(* IEC 61131-3 sources: daoli-st-library/DL_Device (part 30) *)

(* ---- FB_DL_SafetyLightCurtainMute.st ---- *)
// FB_DL_SafetyLightCurtainMute v1.0.0
(*==============================================================================
 * 功能描述: C4 安全光栅消隐。双传感器方向判别消隐状态机：eIdle→eArmed→eMuted→
 *           eRestore→eIdle；双模式下行进方向须 S1 先 S2 后（tDirWin 窗内），方向
 *           错误或消隐超窗 tMuteMax 进 eFault 锁存；单模式下光束遮挡直接进入消隐。
 *           bMuteOut 仅在 eMuted 合法窗口励磁——消隐只放行物料方向判别通过，不屏蔽
 *           任何人体进入判别（muted 不等于屏蔽危险），eFault 相 bMuteOut 强制断磁。
 * 接口契约: 输入 bS1/bS2/bDualMode/bMuteReq/tDirWin/tMuteMax/bReset；
 *           输出 bMuteOut/eState/eCause/bError/nErrId。
 * 边界: ① 组态闸：tDirWin<=T#0S、tMuteMax<=T#0S → 故障锁存；② 三枚 R_TRIG + 两枚
 *           TON 段 0 无条件周期刷新；③ 恢复相再次遮挡判超窗违约（安全侧，不续窗）；
 *           ④ 零全局耦合。
 * 码表: 16#0007_0303 故障级总码（组态非法/方向违约/消隐超窗/非法相位，锁存至 bReset
 *       上升沿且光束全清）；16#0007_0403 信息级：消隐窗口有效（励磁中，每拍重算）。
 * 修订历史: 2026-11-23  v1.0.0  R74 首版
 *==============================================================================*)

TYPE E_DL_SlcState :
(
    eIdle    := 0,    // 待命（光束清、无请求）/ Idle, beams clear, no request
    eArmed   := 10,   // 已布防（等待方向判别）/ Armed, awaiting direction discrimination
    eMuted   := 20,   // 消隐励磁中 / Muted, output energised
    eRestore := 30,   // 恢复相（等待光束全清）/ Restore, awaiting beams clear
    eFault   := 90    // 故障锁存相（复位沿 + 光束全清迁出）/ Fault latched
);
END_TYPE

TYPE E_DL_SlcCause :
(
    eNone       := 0,   // 无故障成因 / No cause
    eCfgIllegal := 1,   // 组态非法 / Illegal configuration
    eDirWrong   := 2,   // 方向判别违约（S2 先于 S1）/ Direction violation, S2 before S1
    eMuteOver   := 3,   // 消隐超窗或恢复相再遮挡 / Mute window overrun or re-break in restore
    ePhaseBad   := 4    // 非法相位兜底 / Illegal phase fallback
);
END_TYPE

FUNCTION_BLOCK FB_DL_SafetyLightCurtainMute
VAR_INPUT
    bS1       : BOOL := FALSE;       // 传感器 1（行进侧首束，TRUE=被遮挡）[-] / Sensor 1, entry side, TRUE = blocked
    bS2       : BOOL := FALSE;       // 传感器 2（行进侧次束，TRUE=被遮挡）[-] / Sensor 2, second beam, TRUE = blocked
    bDualMode : BOOL := TRUE;        // 双传感器方向判别模式（FALSE=单传感器）[-] / Dual-sensor direction mode, FALSE = single
    bMuteReq  : BOOL := FALSE;       // 消隐请求（安全控制器电平）[-] / Mute request from safety controller
    tDirWin   : TIME := T#500MS;     // S1→S2 方向判别窗，域 > T#0S [ms] / Direction window, domain > T#0S
    tMuteMax  : TIME := T#10S;       // 消隐最大励磁窗，域 > T#0S [ms] / Maximum mute window, domain > T#0S
    bReset    : BOOL := FALSE;       // 复位，上升沿清故障锁存 [-] / Reset edge clears fault
END_VAR
VAR_OUTPUT
    bMuteOut  : BOOL;                // 消隐励磁输出（仅合法窗口 TRUE）[-] / Mute output, energised in legal window only
    eState    : E_DL_SlcState;       // 状态出口，段尾单点映射 / State outlet
    eCause    : E_DL_SlcCause;       // 故障成因出口（归因唯一） / Fault cause outlet
    bError    : BOOL;                // 故障锁存标志 [-] / Fault latch flag
    nErrId    : UDINT;               // 事件码，0 = 无事件 / Event code, 0 = none
END_VAR
VAR
    _eState  : E_DL_SlcState := E_DL_SlcState.eIdle;   // 内部相位（CASE 唯一写入目标） / Internal phase
    _eCause  : E_DL_SlcCause := E_DL_SlcCause.eNone;   // 故障成因锁存量 / Latched cause
    rtS1     : R_TRIG;               // S1 上升沿实例，段 0 无条件刷新 / S1 rising edge instance
    rtS2     : R_TRIG;               // S2 上升沿实例，段 0 无条件刷新 / S2 rising edge instance
    rtReset  : R_TRIG;               // 复位沿实例，段 0 无条件刷新 / Reset edge instance
    tonDir   : TON;                  // 方向判别窗计时（S1 遮挡期间），段 0 无条件刷新 / Direction window timer
    tonMute  : TON;                  // 消隐励磁窗计时，段 0 无条件刷新 / Mute window timer
    _bCfgBad : BOOL;                 // 组态非法当拍量 [-] / Illegal configuration this scan
    _bFault  : BOOL;                 // 故障锁存位（锁存量） / Latched fault bit
    _uFault  : UDINT;                // 故障码锁存（锁存量） / Latched fault code
    _uInfo   : UDINT;                // 信息码，每拍重算 / Info code, recomputed each scan
    _bClear  : BOOL;                 // 光束全清当拍量 [-] / All beams clear this scan
    _bArmedOk: BOOL;                 // 布防前置成立当拍量 [-] / Arming precondition this scan
END_VAR

(* —— 段 0：沿实例与定时器无条件周期刷新（禁置于 IF/CASE 内） —— *)
rtS1(CLK := bS1);                                                  // S1 沿，每拍必调 / S1 edge every scan
rtS2(CLK := bS2);                                                  // S2 沿，每拍必调 / S2 edge every scan
rtReset(CLK := bReset);                                            // 复位沿，每拍必调 / Reset edge every scan
tonDir(IN := (_eState = E_DL_SlcState.eArmed) AND bS1, PT := tDirWin);    // 方向窗（布防相 S1 遮挡期）/ Direction timer while armed and S1 blocked
tonMute(IN := (_eState = E_DL_SlcState.eMuted), PT := tMuteMax);   // 消隐窗（励磁相独占）/ Mute timer while muted

(* —— 段 1：单拍量预清零（锁存量 _bFault/_uFault/_eCause 不入清单） —— *)
bError := FALSE;                                                   // 故障标志预清（置位处同拍回填） / Error flag preset
bMuteOut := FALSE;                                                 // 励磁输出预清（eMuted 相回填） / Mute output preset
_uInfo := 16#0000_0000;                                            // 信息码每拍重算 / Info recomputed every scan
nErrId := 16#0000_0000;                                            // 事件码缺省无事件 / Event code default none
_bClear := (NOT bS1) AND (NOT bS2);                                // 光束全清当拍量 / Beams clear this scan
_bArmedOk := _bClear AND bMuteReq AND (NOT _bFault);               // 布防前置：光束清 + 请求在 / Arming precondition

(* —— 段 2：组态域闸 —— *)
_bCfgBad := (tDirWin <= T#0S) OR (tMuteMax <= T#0S);               // 时间域闸（防窗口恒成立） / Time domain gates

(* —— 段 3：故障锁存与解除（R45 配对；解除沿 = 复位沿 + 组态合法 + 光束全清） —— *)
IF _bCfgBad THEN                                                   // 组态非法 / Illegal configuration
    _uFault := 16#0007_0303;                                       // 故障级总码 / Fault-level code
    _bFault := TRUE;
    bError  := TRUE;
    _eCause := E_DL_SlcCause.eCfgIllegal;                          // 归因：组态非法 / Cause: illegal configuration
END_IF
IF rtReset.Q AND (NOT _bCfgBad) AND _bClear THEN                   // 解除沿（当拍量，光束全清） / Release edge with beams clear
    _bFault := FALSE;                                              // 清故障锁存 / Clear fault latch
    _uFault := 16#0000_0000;                                       // 清故障码 / Clear fault code
    _eCause := E_DL_SlcCause.eNone;                                // 清成因 / Clear cause
    IF _eState = E_DL_SlcState.eFault THEN
        _eState := E_DL_SlcState.eIdle;                            // 故障相唯一迁出路径 / Sole exit from fault phase
    END_IF
END_IF

(* —— 段 4：相位机（ENUM 全成员显式标签 + ELSE 兜底） —— *)
CASE _eState OF

E_DL_SlcState.eIdle:
    IF _bFault THEN                                                // 出口 1：故障锁存 / Fault latched
        _eState := E_DL_SlcState.eFault;
    ELSIF _bArmedOk THEN                                           // 出口 2：前置成立进布防 / Preconditions met, arm
        _eState := E_DL_SlcState.eArmed;
    END_IF

E_DL_SlcState.eArmed:
    IF _bFault THEN                                                // 出口 1：故障锁存 / Fault latched
        _eState := E_DL_SlcState.eFault;
    ELSIF (NOT bMuteReq) OR _bCfgBad THEN                          // 出口 2：请求撤销或组态坏 → 回待命 / Request dropped, back to idle
        _eState := E_DL_SlcState.eIdle;
    ELSIF bDualMode THEN                                           // 双传感器模式分支 / Dual-sensor branch
        IF rtS2.Q AND (NOT bS1) THEN                               // 方向违约：S2 先遮挡而 S1 未遮挡 / Direction violation, S2 first
            _uFault := 16#0007_0303;
            _bFault := TRUE;
            bError  := TRUE;
            _eCause := E_DL_SlcCause.eDirWrong;                    // 归因：方向违约 / Cause: direction violation
            _eState := E_DL_SlcState.eFault;
        ELSIF rtS2.Q AND bS1 THEN                                  // 合法方向：S1 已遮挡后 S2 到 → 进励磁 / Legal direction, enter muted
            _eState := E_DL_SlcState.eMuted;
        ELSIF tonDir.Q THEN                                        // S1 遮挡超方向窗（判别失败安全退） / S1 blocked over direction window
            _eState := E_DL_SlcState.eIdle;
        END_IF
    ELSE                                                           // 单传感器模式：遮挡即励磁 / Single mode, block enters muted
        IF bS1 THEN
            _eState := E_DL_SlcState.eMuted;
        END_IF
    END_IF

E_DL_SlcState.eMuted:
    IF _bFault THEN                                                // 出口 1：故障锁存 / Fault latched
        _eState := E_DL_SlcState.eFault;
    ELSIF tonMute.Q THEN                                           // 出口 2：励磁超最大窗 → 强制恢复 / Mute window overrun
        _uFault := 16#0007_0303;                                   // 故障级：消隐超窗（超窗不续磁） / Fault, window overrun
        _bFault := TRUE;
        bError  := TRUE;
        _eCause := E_DL_SlcCause.eMuteOver;                        // 归因：超窗 / Cause: window overrun
        _eState := E_DL_SlcState.eRestore;
    ELSIF (NOT bMuteReq) THEN                                      // 出口 3：请求撤销进恢复 / Request dropped, restore
        _eState := E_DL_SlcState.eRestore;
    ELSE
        _uInfo := 16#0007_0403;                                    // 信息级：消隐励磁中 / Info: mute energised
    END_IF

E_DL_SlcState.eRestore:
    IF _bFault THEN                                                // 出口 1：故障锁存 / Fault latched
        _eState := E_DL_SlcState.eFault;
    ELSIF bS1 OR bS2 THEN                                          // 出口 2：恢复相再遮挡 = 违约（不续窗，安全侧） / Re-break in restore, fault
        _uFault := 16#0007_0303;
        _bFault := TRUE;
        bError  := TRUE;
        _eCause := E_DL_SlcCause.eMuteOver;                        // 归因：恢复相再遮挡 / Cause: re-break in restore
        _eState := E_DL_SlcState.eFault;
    ELSE
        _eState := E_DL_SlcState.eIdle;                            // 出口 3：光束全清回待命 / Beams clear, back to idle
    END_IF

E_DL_SlcState.eFault:
    ;                                                              // 故障相：仅段 3 解除沿可迁出（励磁强制断） / Only the release edge leaves, output forced off

ELSE
    _uFault := 16#0007_0303;                                       // 故障级：非法相位兜底 / Illegal-phase fallback
    _bFault := TRUE;
    bError  := TRUE;
    _eCause := E_DL_SlcCause.ePhaseBad;                            // 归因：非法相位 / Cause: illegal phase
    _eState := E_DL_SlcState.eFault;                               // 强拉故障相 / Force fault phase

END_CASE

(* —— 段 5：出口单点映射（名实同源；锁存码回放；故障相励磁强制断） —— *)
IF (_eState = E_DL_SlcState.eMuted) AND (NOT _bFault) THEN
    bMuteOut := TRUE;                                              // 仅合法励磁相输出 / Output only in legal muted phase
END_IF
IF _bFault THEN
    nErrId := _uFault;                                             // 故障锁存码回放 / Replay latched fault code
ELSE
    nErrId := _uInfo;                                              // 信息码 / Info code
END_IF
bError := _bFault;                                                 // 故障标志与锁存同源 / Flag from latch
eState := _eState;                                                 // 状态出口 / State outlet
eCause := _eCause;                                                 // 成因出口 / Cause outlet

END_FUNCTION_BLOCK

(* ---- FB_DL_SafetyRelayFeedback.st ---- *)
(*==============================================================================
 * 组件名称 (Component)  : FB_DL_SafetyRelayFeedback
 * 所属子库 (Sublibrary) : DL_Device
 * 当前版本 (Version)    : 1.0.0
 * 兼容性   (Platform)   : CODESYS 3.5+ / TwinCAT 3 / 汇川 InoProShop / 施耐德 Machine Expert
 *                         仅依赖 Standard.library（TON / R_TRIG）与库内健康枚举唯一属主，
 *                         零厂商私有库
 * 功能描述 (Function)   : 安全继电器（双通道触点）反馈一致性监视。指令 bCmd 变化后开
 *                         tSyncWin 同步窗，窗内应两通道同步跟随；窗末判定四类结局：
 *                         ① 两通道仍不一致 → 通道不同步故障（eSync）；
 *                         ② 仅通道 1 未跟随 → 通道 1 失效（eCh1Fail）；
 *                         ③ 仅通道 2 未跟随 → 通道 2 失效（eCh2Fail）；
 *                         ④ 两通道都未跟随 → 双通道失效（eBothFail）。
 *                         另连续监视常闭回路断开：bNcLogic 为真时「指令为 FALSE 而两通道反馈
 *                         仍为 FALSE」即常闭回路断开（eNcOpen，典型断线/线圈失电）。
 * 安全声明 (Safety)     : **本件不实现任何安全认证功能**。它是反馈一致性监视器，不是安全功能
 *                         的组成部分：不提供双通道自诊断覆盖率证明，不参与 ISO 13849 / IEC 62061
 *                         的 PL / SIL 定级，其输出不得接入安全链路的停机判据。
 * 归属声明 (Ownership)  : 健康出口 eHealth 引用枚举 `E_DL_Ne107Status` 的**唯一属主**，属主文件为
 *                         `C:\Library\DL_Device\I_DL_DeviceHealth.st`（枚举定义位于该文件 L91 附近），
 *                         本件**只引用不重复声明**（全库同名枚举定义计数必须为 1，R67）。
 * 接口     (Interface)  : 输入 bFbCh1 / bFbCh2 双通道反馈、bCmd 指令、tSyncWin 同步窗、bNcLogic
 *                         常闭逻辑组态位、bReset 复位；输出 eCause 归因、bSyncOk 双通道同步、
 *                         eHealth NE107 健康态、eState / bError / nErrId。
 * 边界     (Boundary)   : ① 组态闸：tSyncWin <= T#0S → 故障锁存，**且非法时 eHealth 直接给
 *                         eFailure**（保守：无法判定同步即按失效上报）；
 *                         ② 常闭语义：bNcLogic = TRUE 时期望反馈 = NOT bCmd；= FALSE 时期望 = bCmd；
 *                         ③ 两通道互斥用布尔 XOR 判，无浮点参与；
 *                         ④ TON 两枚 + R_TRIG 两枚段 0 无条件周期刷新（IN 由相位派生，R228A）；
 *                         ⑤ 故障相迁出唯一路径 = bReset 上升沿；⑥ 零全局耦合（无 GVL / 无物理地址）。
 * 解除式   (Release)    : bReset 上升沿 ∧ 组态合法 ∧ 两通道当前一致（bFbCh1 = bFbCh2，当拍量，
 *                         R240 范式）。自证可满足（终审两式 1）：两枚 TON 的 IN 均挂相位，
 *                         故障相内 IN 恒假 → Q 恒假；两通道物理恢复一致即达，无恒假因子。
 * 码表     (Codes)      : 16#0003_0701 故障级：安全继电器反馈故障总码（组态非法 / 通道不同步 /
 *                         单通道失效 / 双通道失效 / 常闭回路断开 / 非法相位），锁存至 bReset 上升沿，
 *                         归因由 eCause 承载（R190 单件单总码，每个成因成员均有独立赋值点）；
 *                         16#0003_0480 信息级：同步窗正常结束（两通道已按指令同步跟随）。
 *                         加码反证（R90）：同步窗正常结束时 bSyncOk 由假转真，而「一直停在 eRun
 *                         未做过切换」也保持 bSyncOk 为真，二者出口组合无法唯一区分「刚完成一次
 *                         动作确认」与「从未动作」，故立一码留痕。
 *                         码段说明：Device 的 03xx 故障子带已占满（03A0~03FF 连续占位，仅余
 *                         03C5~03C9 碎片孔洞），按实战规则 13「禁止回填他人预留碎片孔洞」，
 *                         本批新开 07xx 故障子带并取 16#0003_0701；信息级仍用 04xx 子带取
 *                         16#0003_0480（该段源码实扫为空）。分段理由即此，非笔误。
 * 开源溯源 (Origin)     : 道莅自研 clean-room（参考 ISA-18.2 / NE107 安全回路一致性语义与
 *                         参数域，零代码行复制；t2-8-isa182 族）
 * 修订历史 (Revision)   : 2026-11-19  v1.0.0  R45 首版（批次 3 · 序号 15）
 *==============================================================================*)

TYPE E_DL_SrfState :
(
    eIdle     := 0,     // 未使能待机 / Idle, standing by
    eSyncWait := 10,    // 指令变化后同步窗内（信号暂不可信） / Inside sync window after a command change
    eRun      := 20,    // 同步完成，稳态监视 / Synchronised, steady monitoring
    eFault    := 90     // 故障锁存相 / Fault latched phase
);
END_TYPE

TYPE E_DL_SrfCause :
(
    eNone       := 0,   // 无故障成因 / No cause
    eCfgIllegal := 1,   // 组态非法 / Illegal configuration
    eSync       := 2,   // 两通道不同步 / Channels out of sync
    eCh1Fail    := 3,   // 通道 1 未跟随 / Channel 1 failed to follow
    eCh2Fail    := 4,   // 通道 2 未跟随 / Channel 2 failed to follow
    eBothFail   := 5,   // 两通道均未跟随 / Both channels failed to follow
    eNcOpen     := 6,   // 常闭回路断开 / Normally-closed loop open
    ePhaseBad   := 7    // 非法相位兜底 / Illegal phase fallback
);
END_TYPE

FUNCTION_BLOCK FB_DL_SafetyRelayFeedback
VAR_INPUT
    bFbCh1    : BOOL := FALSE;          // 通道 1 反馈 [-] / Channel 1 feedback
    bFbCh2    : BOOL := FALSE;          // 通道 2 反馈 [-] / Channel 2 feedback
    bCmd      : BOOL := FALSE;          // 继电器指令 [-] / Relay command
    tSyncWin  : TIME := T#300MS;        // 同步窗时长，域 > T#0S [ms] / Sync window duration, domain > T#0S [ms]
    bNcLogic  : BOOL := TRUE;           // 常闭逻辑组态位：TRUE 时期望反馈 = NOT bCmd [-] / NC logic: expected = NOT command
    bReset    : BOOL := FALSE;          // 复位命令，上升沿清故障 [-] / Reset command, rising edge clears fault
END_VAR
VAR_OUTPUT
    eCause    : E_DL_SrfCause;          // 故障成因出口（R190 归因唯一） / Fault cause outlet
    bSyncOk   : BOOL;                   // 双通道同步（稳态且两通道一致且均符合期望） [-] / Channels in sync
    eHealth   : E_DL_Ne107Status;       // NE107 健康态（引用唯一属主枚举） [-] / NE107 health, owner enum referenced
    eState    : E_DL_SrfState;          // 状态出口，段 6 单点映射 / State outlet
    bError    : BOOL;                   // 故障锁存标志 [-] / Fault latch flag
    nErrId    : UDINT;                  // 事件码，0 = 无事件 / Event code, 0 = no event
END_VAR
VAR
    _eState   : E_DL_SrfState := E_DL_SrfState.eIdle;      // 内部相位（CASE 唯一写入目标） / Internal phase
    _eCause   : E_DL_SrfCause := E_DL_SrfCause.eNone;      // 故障成因锁存（锁存量） / Latched cause
    tonSync   : TON;                    // 同步窗计时，段 0 无条件调用 / Sync window timer
    tonDiff   : TON;                    // 通道不一致持续计时，段 0 无条件调用 / Channel-difference timer
    rtCmd     : R_TRIG;                 // 指令变化沿实例，段 0 无条件调用 / Command change edge
    rtReset   : R_TRIG;                 // 复位沿实例，段 0 无条件调用 / Reset edge
    _bExpect  : BOOL;                   // 常闭/常开语义换算后的期望反馈当拍量 [-] / Expected feedback after NC/NO mapping
    _bChDiff  : BOOL;                   // 两通道不一致当拍量 [-] / Channels disagree
    _bCh1Ok   : BOOL;                   // 通道 1 符合期望当拍量 [-] / Channel 1 matches expectation
    _bCh2Ok   : BOOL;                   // 通道 2 符合期望当拍量 [-] / Channel 2 matches expectation
    _bNcOpen  : BOOL;                   // 常闭回路断开当拍量 [-] / NC loop open
    _bCfgBad  : BOOL;                   // 组态非法当拍量 [-] / Illegal configuration
    _bFault   : BOOL;                   // 故障锁存位（锁存量） / Latched fault bit
    _uFault   : UDINT;                  // 故障码锁存（锁存量） / Latched fault code
    _uInfo    : UDINT;                  // 信息码，每拍重算 / Info code, recomputed each scan
END_VAR

(* —— 段 0：当拍判据派生 + 定时器与沿实例无条件周期刷新 —— *)
_bExpect := bCmd;                                                                  // 缺省常开语义 / Default NO logic
IF bNcLogic THEN
    _bExpect := NOT bCmd;                                                          // 常闭语义：期望反馈取反 / NC logic inverts the expectation
END_IF
_bChDiff := bFbCh1 XOR bFbCh2;                                                     // 两通道不一致（布尔异或） / Channels disagree
_bCh1Ok  := (bFbCh1 AND _bExpect) OR ((NOT bFbCh1) AND (NOT _bExpect));             // 通道 1 符合期望 / Channel 1 matches expectation
_bCh2Ok  := (bFbCh2 AND _bExpect) OR ((NOT bFbCh2) AND (NOT _bExpect));             // 通道 2 符合期望 / Channel 2 matches expectation
_bNcOpen := bNcLogic AND (NOT bCmd) AND (NOT bFbCh1) AND (NOT bFbCh2);              // 常闭回路断开（指令 0 而反馈 0） / NC loop open
_bCfgBad := (tSyncWin <= T#0S);                                                     // 组态域闸 / Configuration gate
rtCmd(CLK := bCmd);                                                                 // 指令变化沿，每拍必调（R228A） / Command change edge
rtReset(CLK := bReset);                                                             // 复位沿，每拍必调 / Reset edge
tonSync(IN := (_eState = E_DL_SrfState.eSyncWait), PT := tSyncWin);                 // 同步窗计时（IN 由相位派生） / Sync window timer
tonDiff(IN := (_eState = E_DL_SrfState.eSyncWait) AND _bChDiff, PT := tSyncWin);    // 不一致持续计时 / Channel-difference timer

(* —— 段 1：单拍量预清零（锁存量不入清单，R107） —— *)
_uInfo   := 16#0000_0000;          // 信息码每拍重算 / Info recomputed every scan
bSyncOk  := FALSE;                 // 同步位每拍预清 / Sync flag preset
nErrId   := 16#0000_0000;          // 事件码缺省无事件 / Event code default none
bError   := FALSE;                 // 故障标志每拍预清，故障分支同拍置位（R45 配对） / Flag preset

(* —— 段 2：复位沿 + 组态域闸 + 常闭断开判决 —— *)
IF rtReset.Q THEN                                                        // 当拍复位沿 / current-scan reset edge
    _bFault := FALSE;                                                    // 清故障锁存位（锁存量） / Clear fault latch
    _uFault := 16#0000_0000;                                             // 清故障锁存码（锁存量） / Clear latched code
    _eCause := E_DL_SrfCause.eNone;                                      // 清成因（锁存量） / Clear latched cause
    IF _eState = E_DL_SrfState.eFault THEN
        _eState := E_DL_SrfState.eIdle;                                  // 故障相迁出唯一路径 / Sole exit from fault phase
    END_IF
END_IF
IF _bCfgBad THEN                                                         // 组态域闸 / Configuration gate
    _uFault := 16#0003_0701;                                             // 故障级：安全继电器反馈故障总码 / Fault-level: relay feedback fault code
    _bFault := TRUE;
    bError  := TRUE;                                                     // 故障标志同拍置位（R45 配对） / Error flag set same scan
    _eCause := E_DL_SrfCause.eCfgIllegal;                                // 归因：组态非法 / Cause: illegal configuration
END_IF
IF (NOT _bFault) AND _bNcOpen THEN                                       // 常闭回路断开（连续监视，不限相位） / NC loop open, monitored continuously
    _uFault := 16#0003_0701;
    _bFault := TRUE;
    bError  := TRUE;
    _eCause := E_DL_SrfCause.eNcOpen;                                    // 归因：常闭断开 / Cause: NC loop open
END_IF

(* —— 段 3：同步窗末判定（四结局归因唯一，R190） —— *)
IF (NOT _bFault) AND tonSync.Q THEN                                      // 同步窗到时 / Sync window elapsed
    IF _bChDiff THEN                                                     // 结局 1：两通道仍不一致 / Outcome 1, still disagreeing
        _uFault := 16#0003_0701;
        _bFault := TRUE;
        bError  := TRUE;
        _eCause := E_DL_SrfCause.eSync;                                  // 归因：不同步 / Cause: out of sync
    ELSIF (NOT _bCh1Ok) AND (NOT _bCh2Ok) THEN                           // 结局 2：两通道均未跟随 / Outcome 2, both failed
        _uFault := 16#0003_0701;
        _bFault := TRUE;
        bError  := TRUE;
        _eCause := E_DL_SrfCause.eBothFail;                              // 归因：双通道失效 / Cause: both channels failed
    ELSIF NOT _bCh1Ok THEN                                               // 结局 3：仅通道 1 未跟随 / Outcome 3, channel 1 only
        _uFault := 16#0003_0701;
        _bFault := TRUE;
        bError  := TRUE;
        _eCause := E_DL_SrfCause.eCh1Fail;                               // 归因：通道 1 失效 / Cause: channel 1 failed
    ELSIF NOT _bCh2Ok THEN                                               // 结局 4：仅通道 2 未跟随 / Outcome 4, channel 2 only
        _uFault := 16#0003_0701;
        _bFault := TRUE;
        bError  := TRUE;
        _eCause := E_DL_SrfCause.eCh2Fail;                               // 归因：通道 2 失效 / Cause: channel 2 failed
    ELSE
        _uInfo := 16#0003_0480;                                          // 信息级：同步窗正常结束 / Info: sync window closed normally
    END_IF
END_IF

(* —— 段 4：故障解除式（R240 全当拍量） —— *)
IF rtReset.Q AND (NOT _bCfgBad) AND (NOT _bChDiff) THEN
    _bFault := FALSE;                                                    // 清故障锁存位（锁存量） / Clear fault latch
    _uFault := 16#0000_0000;                                             // 清故障锁存码（锁存量） / Clear latched code
    _eCause := E_DL_SrfCause.eNone;                                      // 清成因（锁存量） / Clear latched cause
END_IF

(* —— 段 4A：故障锁存相位迁移闸 —— *)
IF _bFault AND (_eState <> E_DL_SrfState.eFault) THEN
    _eState := E_DL_SrfState.eFault;                                     // 锁存即入故障相 / Latch enters fault phase
END_IF

(* —— 段 5：相位机（ENUM 全成员显式标签 + ELSE 兜底，R128） —— *)
CASE _eState OF

E_DL_SrfState.eIdle:
    IF (NOT _bCfgBad) AND (NOT _bFault) THEN                             // 出口 1：组态合法，进入稳态监视 / Config legal, enter steady monitoring
        _eState := E_DL_SrfState.eRun;
    ELSIF _bFault THEN                                                   // 出口 2：故障锁存 / Fault latched
        _eState := E_DL_SrfState.eFault;
    END_IF

E_DL_SrfState.eRun:
    IF rtCmd.Q AND (NOT _bFault) THEN                                    // 出口 1：指令变化，开同步窗 / Command changed, open sync window
        _eState := E_DL_SrfState.eSyncWait;
    ELSIF _bFault THEN                                                   // 出口 2：故障锁存 / Fault latched
        _eState := E_DL_SrfState.eFault;
    END_IF

E_DL_SrfState.eSyncWait:
    IF tonSync.Q THEN                                                    // 出口 1：窗到，判定已由段 3 完成 / Window elapsed, verdict done in segment 3
        IF _bFault THEN
            _eState := E_DL_SrfState.eFault;                             // 判定失败即入故障相 / Failed verdict enters fault
        ELSE
            _eState := E_DL_SrfState.eRun;                               // 同步成功回稳态 / Sync OK back to steady run
        END_IF
    ELSIF (NOT bCmd) AND (NOT _bChDiff) THEN                             // 出口 2：指令回安全侧且两通道已一致（判据对象消失，R98） / Command back on the safe side with channels consistent
        _eState := E_DL_SrfState.eRun;
    END_IF

E_DL_SrfState.eFault:
    ;                                                                     // 故障相：仅段 4 复位沿可迁出 / Only the reset edge leaves this phase

ELSE
    _uFault := 16#0003_0701;                                             // 故障级：非法相位兜底（归并总码） / Illegal-phase fallback
    _bFault := TRUE;
    bError  := TRUE;
    _eCause := E_DL_SrfCause.ePhaseBad;                                  // 归因：非法相位 / Cause: illegal phase
    _eState := E_DL_SrfState.eFault;

END_CASE

(* —— 段 6：出口单点映射（名实同源；锁存码回放；NE107 健康态仲裁） —— *)
IF _bFault OR _bCfgBad THEN
    bSyncOk := FALSE;                                                    // 故障/组态非法：不宣称同步 / No sync claim
    eHealth := E_DL_Ne107Status.eFailure;                                // 失效级（组态非法也按失效保守上报） / Failure level, conservative
ELSIF _eState = E_DL_SrfState.eSyncWait THEN
    bSyncOk := FALSE;                                                    // 窗内信号暂不可信 / Signals not yet trustworthy inside the window
    eHealth := E_DL_Ne107Status.eCheckFunction;                          // 功能检查级：动作确认中 / Function-check level during confirmation
ELSIF (_eState = E_DL_SrfState.eRun) AND (NOT _bChDiff) AND _bCh1Ok AND _bCh2Ok THEN
    bSyncOk := TRUE;                                                     // 稳态且两通道一致且符合期望 / Steady, consistent and as expected
    eHealth := E_DL_Ne107Status.eOk;                                     // 正常级 / OK level
ELSE
    bSyncOk := FALSE;                                                    // 其余情形一律不宣称同步 / No sync claim otherwise
    eHealth := E_DL_Ne107Status.eMaintenanceReq;                         // 需要维护级 / Maintenance-required level
END_IF
IF _bFault THEN
    nErrId := _uFault;                                                   // 故障锁存码回放 / Replay latched fault code
ELSE
    nErrId := _uInfo;                                                    // 信息码 / Info code
END_IF
bError := _bFault;                                                       // 故障标志与锁存同源（名实双出口，R191） / Flag from latch
eState := _eState;                                                       // 状态出口 / State outlet
eCause := _eCause;                                                       // 成因出口 / Cause outlet

END_FUNCTION_BLOCK

(* ---- FB_DL_SealIntegrityMonitor.st ---- *)
(*==============================================================================
 * 组件名称 (Component)  : FB_DL_SealIntegrityMonitor
 * 所属子库 (Sublibrary) : DL_Device
 * 当前版本 (Version)    : 1.0.0
 * 兼容性 (Platform)     : CODESYS 3.5 / TwinCAT 3 / 汇川 InoProShop / Machine Expert
 *                         仅依赖纯 IEC 61131-3 标准元素，零厂商方言
 * 功能描述 (Function)   : 封口完整性在线监视（仅监视不执行封口）：bSealDone
 *                         上升沿采样温度/压力/时间三值，与配方窗独立比对，全过
 *                         → bInSpec；NaN 判超差；连续超差计数达阈值 → 预警锁存
 *                         （需复位）；窗下限 < 上限合法性自检，非法拒绝判定。
 * 溯源 (Origin)         : 道莅 clean-room 防御性实现
 * 本文件内含 (Contains) : TYPE E_DL_SealErr / FUNCTION_BLOCK FB_DL_SealIntegrityMonitor
 * 依赖 (Depends)        : 无 DL_ 内部依赖；Standard.library R_TRIG 实例
 * 红线自检 (Redline)    : 无外部全局变量、无硬件地址直引 ｜ 全变量中英双语同行注释
 *                         窗参数合法性自检 ｜ NaN 判超差 ｜ 计数饱和 65535 ｜
 *                         枚举成员全部显式赋值 ｜ R_TRIG 实例每周期无条件调用 ｜
 *                         主码取首个违参（温度 > 压力 > 时间优先级）禁浮点判等
 * 错误码表 (Codes)      : 16#0003_03A2 在规格内
 *                         16#0003_03A3 温度超差
 *                         16#0003_03A4 压力超差
 *                         16#0003_03A5 时间超差
 *                         16#0003_03A6 故障级 窗参数非法(拒绝判定)
 * 修订历史 (Revision)   : 2026-11-17  v1.0.0  首版入库 · R27 · 阶段三批 2
 * 验收向量 (Acceptance) : 窗 180~220 C / 300~400 N / T#800MS~T#1200MS：
 *                         三值 200/350/1000ms → 03A2；温度 230 → 03A3 连续 3 次 → 预警锁存
 *============================================================================*)

(*-----------------------------------------------------------------------------
 * 枚举: E_DL_SealErr（归属 DL_Device，与 FB_DL_SealIntegrityMonitor 同文件）
 *----------------------------------------------------------------------------*)
TYPE E_DL_SealErr :
(
    eInSpec     := 16#0003_03A2,   // 在规格内 / Within specification
    eTempViol   := 16#0003_03A3,   // 温度超差 / Temperature violation
    ePressViol  := 16#0003_03A4,   // 压力超差 / Pressure violation
    eTimeViol   := 16#0003_03A5,   // 时间超差 / Time violation
    eWindowBad  := 16#0003_03A6    // 故障级：窗参数非法，拒绝判定 / Fault: illegal window, judging refused
);
END_TYPE

(*==============================================================================
 * 功能块: FB_DL_SealIntegrityMonitor
 * 调用约定: 每个扫描周期无条件调用一次。
 *============================================================================*)
FUNCTION_BLOCK FB_DL_SealIntegrityMonitor
VAR_INPUT
    fSealTemp_C  : REAL;               // 封口温度 [摄氏度] / Seal temperature [degC]
    fSealPress_N : REAL;               // 封口压力 [牛] / Seal pressure [N]
    tSealTime    : TIME;               // 封口时间 [毫秒] / Seal time [ms]
    fTempWin_L   : REAL;               // 温度窗下限 [摄氏度] / Temperature window low [degC]
    fTempWin_H   : REAL;               // 温度窗上限 [摄氏度] / Temperature window high [degC]
    fPressWin_L  : REAL;               // 压力窗下限 [牛] / Pressure window low [N]
    fPressWin_H  : REAL;               // 压力窗上限 [牛] / Pressure window high [N]
    tTimeWin_L   : TIME;               // 时间窗下限 [毫秒] / Time window low [ms]
    tTimeWin_H   : TIME;               // 时间窗上限 [毫秒] / Time window high [ms]
    uViolTrip    : UINT := 3;          // 连续超差预警阈值 [次] / Consecutive-violation trip threshold [pcs]
    bSealDone    : BOOL;               // 封口节拍完成（上升沿采样）/ Seal cycle done, sampled on rising edge
    bReset       : BOOL;               // 预警锁存复位 / Alarm latch reset
END_VAR
VAR_OUTPUT
    bInSpec      : BOOL;               // 三参全在窗内 / All three parameters in window
    bAlarmLatch  : BOOL;               // 预警锁存（连续超差达阈值）/ Alarm latch, threshold reached
    nViolCnt     : UINT;               // 连续超差次数 [次] / Consecutive violation count [pcs]
    eError       : E_DL_SealErr;       // 主错误码（取首个违参）/ Main error code, first violated parameter
END_VAR
VAR
    fbSealTrig   : R_TRIG;             // 封口节拍上升沿实例（无条件调用）/ Seal-done edge instance
    fbResetTrig  : R_TRIG;             // 复位上升沿实例（无条件调用）/ Reset edge instance
    bTempOk      : BOOL;               // 温度窗内判据 / Temperature in-window predicate
    bPressOk     : BOOL;               // 压力窗内判据 / Pressure in-window predicate
    bTimeOk      : BOOL;               // 时间窗内判据 / Time in-window predicate
    bWindowOk    : BOOL;               // 窗参数合法性判据 / Window legality predicate
    bTempValid   : BOOL;               // 温度非有限有效 / Temperature finite validity
    bPressValid  : BOOL;               // 压力非有限有效 / Pressure finite validity
    uViolTripUse : UINT;               // 生效预警阈值（下限钳 1）[次] / Effective trip threshold [pcs]
END_VAR
VAR CONSTANT
    DL_SEAL_INF_MAX  : REAL := 1.0E30;      // 非有限值判定幅值上限 / Magnitude bound for finite-value check
    DL_SEAL_CNT_SAT  : UINT := 65535;       // 超差计数饱和值 [次] / Violation count saturation [pcs]
    DL_SEAL_TRIP_MIN : UINT := 1;           // 预警阈值下限 [次] / Trip threshold lower bound [pcs]
END_VAR

(*------------------------------------------------------------------------------
 * 段 1｜R_TRIG 实例每周期无条件调用（仅输入条件化）
 *----------------------------------------------------------------------------*)
fbSealTrig(CLK := bSealDone);                        // 封口节拍沿检测无条件刷新 / seal edge refreshed unconditionally
fbResetTrig(CLK := bReset);                          // 复位沿检测无条件刷新 / reset edge refreshed unconditionally

(*------------------------------------------------------------------------------
 * 段 2｜窗参数合法性自检：下限必须严格小于上限，非法则拒绝判定（故障级）
 *----------------------------------------------------------------------------*)
bWindowOk := (fTempWin_L < fTempWin_H) AND (fPressWin_L < fPressWin_H) AND (tTimeWin_L < tTimeWin_H);   // 三窗合法性 / three-window legality
IF NOT bWindowOk THEN
    eError := E_DL_SealErr.eWindowBad;               // 故障级：窗参数非法 / fault: illegal window
    bInSpec := FALSE;                                // 拒绝判定：规格输出 FALSE / judging refused
    nViolCnt := 0;                                   // 计数清零（非法窗不计超差）/ count cleared
    RETURN;
END_IF

(*------------------------------------------------------------------------------
 * 段 3｜阈值下限钳位与复位沿处理
 *----------------------------------------------------------------------------*)
uViolTripUse := uViolTrip;                           // 阈值工作副本 / threshold working copy
IF uViolTripUse < DL_SEAL_TRIP_MIN THEN
    uViolTripUse := DL_SEAL_TRIP_MIN;                // 阈值下限钳位 / threshold floored
END_IF
IF fbResetTrig.Q THEN
    bAlarmLatch := FALSE;                            // 复位解锁存 / unlatch on reset
    nViolCnt := 0;                                   // 计数清零 / count cleared
END_IF

(*------------------------------------------------------------------------------
 * 段 4｜节拍采样判定（bSealDone 上升沿一次性判定，非沿拍保持上拍结果）
 *----------------------------------------------------------------------------*)
IF fbSealTrig.Q THEN
    bTempValid := (fSealTemp_C = fSealTemp_C) AND (ABS(fSealTemp_C) <= DL_SEAL_INF_MAX);   // 温度非有限有效 / temperature finite
    bPressValid := (fSealPress_N = fSealPress_N) AND (ABS(fSealPress_N) <= DL_SEAL_INF_MAX);   // 压力非有限有效 / pressure finite
    bTempOk := bTempValid AND (fSealTemp_C >= fTempWin_L) AND (fSealTemp_C <= fTempWin_H);   // 温度窗内（NaN 判超差）/ temp in window
    bPressOk := bPressValid AND (fSealPress_N >= fPressWin_L) AND (fSealPress_N <= fPressWin_H);   // 压力窗内 / pressure in window
    bTimeOk := (tSealTime >= tTimeWin_L) AND (tSealTime <= tTimeWin_H);   // 时间窗内 / time in window
    bInSpec := bTempOk AND bPressOk AND bTimeOk;     // 三参全在窗 / all in window
    IF bInSpec THEN
        nViolCnt := 0;                               // 合格清连续计数 / clear consecutive count
        eError := E_DL_SealErr.eInSpec;              // 码 03A2 / code in-spec
    ELSE
        IF nViolCnt < DL_SEAL_CNT_SAT THEN
            nViolCnt := nViolCnt + 1;                // 连续超差计数饱和自增 [次] / saturating violation increment
        END_IF
        IF bTempOk THEN
            eError := E_DL_SealErr.ePressViol;       // 温度合格则主码取压力（首个违参优先级压力次之）/ main code picks pressure
        ELSIF bPressOk THEN
            eError := E_DL_SealErr.eTimeViol;        // 压力合格则主码取时间 / main code picks time
        ELSE
            eError := E_DL_SealErr.eTempViol;        // 温度违参优先取主码（首个违参 = 温度最优先）/ main code picks temperature first
        END_IF
        IF nViolCnt >= uViolTripUse THEN
            bAlarmLatch := TRUE;                     // 连续超差达阈值：预警锁存 / threshold reached: alarm latched
        END_IF
    END_IF
END_IF
END_FUNCTION_BLOCK

(* ---- FB_DL_SensorGlitchFilter.st ---- *)
// FB_DL_SensorGlitchFilter v1.0.0
// 开源溯源：来源 brOscatLib / URL https://github.com/iec-oscat-mirror / 许可证 MIT / 借鉴点 FT_IMP 一阶惯性滤波语义
(*==============================================================================
 * 功能描述: 传感器毛刺滤波单件。|Δ| > fGlitchBand 计为疑似毛刺并计数，连续超
 *           nFollowCnt 拍才跟随（真实阶跃），否则保持上一拍值并置 bGlitch；正常域
 *           内以一阶惯性 fAlpha 平滑跟随。非有限输入防御（保持 + bValid=FALSE），
 *           组态非法（带宽/惯性系数/计数域）防御。
 * 接口契约: 输入 fRaw/fGlitchBand/nFollowCnt/fAlpha/bEnable；
 *           输出 fFiltered/bValid/bGlitch。
 * 边界: 零定时器零沿实例（纯逐拍滤波），零全局耦合；bEnable=FALSE 时输出冻结保持。
 * 修订历史: 2026-11-23  v1.0.0  R74 首版
 *==============================================================================*)

FUNCTION_BLOCK FB_DL_SensorGlitchFilter
VAR_INPUT
    fRaw        : REAL := 0.0;     // 原始采样输入 [工程单位] / Raw sample input
    fGlitchBand : REAL := 1.0;     // 毛刺判别带宽，域 > 0 [工程单位/拍] / Glitch band [unit/scan]
    nFollowCnt  : INT := 3;        // 疑似毛刺连续计数门槛（超 N 拍才跟随）[拍] / Consecutive count threshold [scan]
    fAlpha      : REAL := 0.2;     // 一阶惯性平滑系数，域 (0,1] [-] / First-order smoothing factor
    bEnable     : BOOL := TRUE;    // 使能（FALSE 输出冻结保持）[-] / Enable, FALSE freezes output
END_VAR
VAR_OUTPUT
    fFiltered : REAL := 0.0;       // 滤波输出 [工程单位] / Filtered output
    bValid    : BOOL;              // 输出有效回执（首拍后为真）[-] / Output validity receipt
    bGlitch   : BOOL;              // 本拍毛刺判别标志（未跟随即真）[-] / Glitch flag this scan
END_VAR
VAR
    _fLast  : REAL := 0.0;         // 上一拍跟随值（锁存量）[工程单位] / Last followed value
    _nCnt   : INT := 0;            // 疑似毛刺连续计数（锁存量）[拍] / Consecutive glitch count
    _bInit  : BOOL := FALSE;       // 首拍初始化标志（锁存量） / First-scan init flag
    _fDelta : REAL := 0.0;         // 本拍增量 [工程单位] / Increment this scan
    _bCfgBad: BOOL;                // 组态非法当拍量 [-] / Illegal configuration this scan
    _bNonFin: BOOL;                // 输入非有限当拍量 [-] / Non-finite input this scan
END_VAR

(* —— 段 0：单拍量预清零（锁存量 _fLast/_nCnt/_bInit 不入清单） —— *)
bValid := FALSE;                             // 有效回执预清 / Validity preset
bGlitch := FALSE;                            // 毛刺标志预清 / Glitch preset

(* —— 段 1：组态域闸与非有限闸（覆盖全部参与引脚） —— *)
_bCfgBad := (fGlitchBand <= 0.0) OR (fGlitchBand <> fGlitchBand)   // 带宽域与 NaN 闸 / Band domain and NaN gate
         OR (nFollowCnt < 1)                            // 计数域闸 / Count domain gate
         OR (fAlpha <= 0.0) OR (fAlpha > 1.0) OR (fAlpha <> fAlpha);   // 惯性系数域与 NaN 闸 / Alpha domain and NaN gate
_bNonFin := fRaw <> fRaw;                    // 输入 NaN 自反判 / Input NaN test

(* —— 段 2：滤波主体（首拍直取；毛刺判别 → 计数 → 跟随/保持；全部逐拍无状态残留） —— *)
IF (NOT bEnable) OR _bCfgBad OR _bNonFin THEN   // 非使能/组态坏/非有限：输出冻结保持 / Frozen hold paths
    IF _bNonFin THEN                         // 非有限输入明确不宣称有效 / Non-finite invalidates receipt
        bValid := FALSE;
    ELSE
        bValid := _bInit;                    // 冻结保持沿用首拍后有效性 / Frozen hold keeps receipt
    END_IF
ELSIF NOT _bInit THEN                        // 首拍：直取输入建立基线 / First scan seeds the baseline
    _fLast := fRaw;                          // 基线装载 / Baseline seeded
    _bInit := TRUE;                          // 首拍完成 / First scan done
    _nCnt := 0;                              // 计数清零 / Count cleared
    fFiltered := _fLast;                     // 输出首拍值 / Output first value
    bValid := TRUE;                          // 有效回执 / Validity receipt
ELSE
    _fDelta := fRaw - _fLast;                // 本拍增量 [工程单位] / Increment this scan
    IF ABS(_fDelta) > fGlitchBand THEN       // 超带宽疑似毛刺 / Over band, suspected glitch
        IF _nCnt < 32000 THEN _nCnt := _nCnt + 1; END_IF   // 连续计数递增（饱和钳位防 INT 回绕） / Count up with saturation clamp
        IF _nCnt >= nFollowCnt THEN          // 连续超 N 拍 → 判真实阶跃，跟随 / Real step, follow
            _fLast := fRaw;                  // 跟随装载 / Follow the input
            _nCnt := 0;                      // 计数归零 / Count reset
            fFiltered := _fLast;             // 输出跟随值 / Output follows
            bGlitch := FALSE;                // 非毛刺（已确认为阶跃） / Not a glitch anymore
        ELSE
            bGlitch := TRUE;                 // 未达计数 → 保持并报毛刺 / Hold and flag glitch
            fFiltered := _fLast;             // 输出保持上一拍 / Output holds last
        END_IF
    ELSE
        _nCnt := 0;                          // 带宽内计数归零 / Within band, count reset
        _fLast := _fLast + fAlpha * (fRaw - _fLast);   // 一阶惯性平滑跟随 / First-order smoothing follow
        fFiltered := _fLast;                 // 输出平滑值 / Output smoothed value
    END_IF
    bValid := TRUE;                          // 有效回执 / Validity receipt
END_IF

END_FUNCTION_BLOCK

(* ---- FB_DL_SensorPairPlausibility.st ---- *)
(*
  ==================================================================
  组件名 Component  : FB_DL_SensorPairPlausibility
  分类   Category   : DL_Device
  前缀   Naming     : FB_DL_ ｜ b/n/u/f/t/e/st 类型前缀制（R265）
  复杂度 Complexity  : 高
  版本   Version    : 1.0.1
  功能   Purpose    : 双冗余传感器交叉合理性（偏差窗 + 漂移趋势 + 择优输出 + 故障锁定状态机）。
  来源   Source     : t2-6-rockwell-aoi（冗余交叉判据公开语义）
  平台   Platform   : 纯 IEC 61131-3（TON 无 / R_TRIG / CASE / FOR），三平台通用
  分工声明 Split     : 与 FB_DL_SensorDriftBaseline（基线学习属主）分工——后者
                      学慢漂基线；本件做双冗余交叉判与择优（R216 双向互引）。
  作者   Author     : 道莅代码库 · PLC 编程专家（R61）
  归属 Ownership     : E_DL_SensorPairPhase 属主为本文件（全库唯一定义，R264）；
                      引用件只引用不重声明。
  ------------------------------------------------------------------
  边界 Boundary     :
                      一 择优切换须迟滞：源切换仅在「当前源非有限」时发生（有效性
                         边界迟滞），合法但分歧时不拍拍翻转（防抖动纪律）；切换
                         拍发单拍 bSwitched（R256 统一出口预置）；
                      二 偏差窗与漂移趋势滚动窗长度 nTrendWin 提为输入（合法域
                         1..32，越域钳位信息级 070A）；窗长变更沿（_nUse ≠ _nUsePrev）
                         全窗清零（和 / 写头 / 填充计数 / 环元素逐项清），防窗长缩小后
                         旧条目永久留在和里（v1.0.1 修 D4 环窗残留）；
                      三 非有限闸逐个点名 fA / fB / fDevWin / fDriftLim 四个浮点
                         入参（R272 全量枚举）；
                      四 故障锁存逐条自证：双传感器偏差超窗（0707）与漂移趋势
                         超限（0708）独立锁存独立码（R190），bReset 上升沿解除
                         （恒可达，R152 自证）；故障相输出冻结最近有效择优快照
                         （R273 快照防污染：快照写前过有限闸）；
                      五 CASE 必带 ELSE 兜底；R_TRIG 段 0 无条件刷新；
                      六 无全局、无外部变量、无物理地址。
  错误码   Codes    :
    16#0003_0707【故障级】双传感器偏差超窗，输出冻结快照，锁存至复位沿
    16#0003_0708【故障级】漂移趋势超限，输出冻结快照，锁存至复位沿
    16#0003_0709【信息级】发生择优源切换（bSwitched 同拍置位）
    16#0003_070A【信息级】滚动窗长度越域已钳位（1..32）
  验收   Acceptance :
    算法已证（脚本）：未跑 ｜ 编译器已证（三平台）：未跑
    V1 A=100/B=100.5、窗 2.0 → fSel=100（A 源）、无故障
    V2 A=NaN → 切 B 源、码 0709、bSwitched 单拍
    V3 B=110（窗 2.0）持续 → 码 0707、输出冻结快照、锁存待复位
    V4 窗 32 跑 40 拍后缩到 8 → 均值只含最近 8 个样本（旧版含陈旧项；v1.0.1 回归）
    V5 窗 8 首 3 拍（_nFill=3）→ 均值 = 3 样本均值（旧版除子 8，偏小 62%）
    V6 双源均非有限（_nFill=0 路径）→ 判据不执行、无除零、无锁存
    V7 窗长 8↔32 反复抖动 → 无残留累加漂移（环元素随变更沿清零）
  修订记录 Revision  :
    2026-11-21  v1.0.0  R61 首版（批 4 · 序号 13）
    2026-11-21  v1.0.1  R62-D4 返修：①新增 _nUsePrev，窗长变更沿全窗清零（含环元素逐项清，防减项把陈旧样本重新注入和）；②新增 _nFill，均值除子由 _nUse 改为 _nFill（首填偏小防漏报）；③_nFill=0 跳过判据并重写除子 ≥1 证明注释；④复位清单补 _nFill / _nUsePrev。注：盘面实测入库版本为 v1.0.0（计划书假设 R61 已发 v1.0.1），按实测优先、禁跳号递增一次至 v1.0.1
  ==================================================================
*)
TYPE E_DL_SensorPairPhase :
(
    eUseA   := 0,  // 择优 A 源 / using the source A
    eUseB   := 10, // 择优 B 源 / using the source B
    eFault  := 20  // 故障锁定：输出冻结快照 / fault locked, the outlet frozen at the snapshot
);
END_TYPE

FUNCTION_BLOCK FB_DL_SensorPairPlausibility
VAR_INPUT
    bEnable   : BOOL := TRUE;   // 使能，FALSE 时冻结择优出口（R191 声明行）/ the enable, false freezes the outlet
    bReset    : BOOL := FALSE;  // 故障复位电平，上升沿清锁存 / the fault reset level
    fA        : LREAL := 0.0;   // A 传感器测量值 [工程单位] / the sensor A value
    fB        : LREAL := 0.0;   // B 传感器测量值 [工程单位] / the sensor B value
    fDevWin   : LREAL := 2.0;   // 偏差窗 [工程单位]，必须 > 0 / the deviation window, must be positive
    fDriftLim : LREAL := 5.0;   // 漂移趋势限 [工程单位]，必须 > 0 / the drift trend limit, must be positive
    nTrendWin : DINT  := 8;     // 漂移趋势滚动窗长度 [拍]，合法域 1..32 / the rolling window length, legal from one to thirty two
END_VAR
VAR_OUTPUT
    fSel      : LREAL := 0.0;  // 择优输出 [工程单位] / the selected outlet
    bSrcA     : BOOL := TRUE;  // 当前择优 A 源指示 [-] / the source A indicator
    bSrcB     : BOOL := FALSE; // 当前择优 B 源指示 [-] / the source B indicator
    bSwitched : BOOL := FALSE; // 源切换单拍脉冲 [-] / the source switch one shot pulse
    eState    : E_DL_SensorPairPhase; // 主状态机当前态 [状态] / the current state
    bError    : BOOL := FALSE; // 故障锁存位（与锁存同源，R191）/ the fault bit from the latch
    bValid    : BOOL := FALSE; // 择优可用标志 [-] / the selection usable flag
    eErr      : UDINT := 16#0000_0000; // 错误码，0 = 正常 / the error code, zero is ok
END_VAR
VAR
    _bInit    : BOOL := FALSE;                          // 首拍初始化标志（R310）/ the first scan flag
    _eState   : E_DL_SensorPairPhase := E_DL_SensorPairPhase.eUseA; // 内部状态寄存器 / the internal state register
    _bFault   : BOOL := FALSE;                          // 故障锁存副本（仅复位沿清除）/ the fault latch copy
    _bDevFlt  : BOOL := FALSE;                          // 偏差超窗锁存副本（独立成因，R190）/ the deviation fault latch copy
    _bDriftFlt: BOOL := FALSE;                          // 漂移超限锁存副本（独立成因）/ the drift fault latch copy
    _bFin     : BOOL := FALSE;                          // 入参非有限闸结果（逐拍重算）/ the finiteness gate result
    _bFinA    : BOOL := FALSE;                          // A 源有限标记（逐拍重算）/ the A finiteness flag
    _bFinB    : BOOL := FALSE;                          // B 源有限标记 / the B finiteness flag
    _fDev     : LREAL := 0.0;                           // 本拍偏差 [工程单位] / the deviation this scan
    _fSnap    : LREAL := 0.0;                           // 最近有效择优快照（写前过闸，FB32-7）/ the last valid snapshot gated before write
    _nUse     : DINT := 8;                              // 钳位后的滚动窗长度 [拍] / the clamped window length
    _afRing   : ARRAY[0..31] OF LREAL;                  // 偏差滚动环形窗 [工程单位] / the deviation rolling ring
    _nHead    : DINT := 0;                              // 环形窗写头 [下标] / the ring write head
    _nFill    : DINT := 0;                              // 环形窗已填样本数 [拍]，均值除子（v1.0.1 修 D4）/ the filled sample count of the ring, the mean divisor
    _nUsePrev : DINT := 0;                              // 上拍窗长快照 [拍]，置 0 使首拍必触发一次全窗清零 / the previous window length snapshot, zero forces a full clear on the first scan
    _nRingIdx : DINT := 0;                              // 环元素清零遍历索引 [下标] / the ring clearing traversal index
    _fRingSum : LREAL := 0.0;                           // 环窗偏差和 [工程单位] / the ring deviation sum
    _bSw      : BOOL := FALSE;                          // 切换单拍内部位，段 1 预清段 5 映射 / the internal switch bit
    _bWinBad  : BOOL := FALSE;                          // 窗长钳位标记（逐拍重算）/ the window clamp flag
    rtReset   : R_TRIG; // 复位沿实例，段 0 无条件刷新 / the reset edge instance
END_VAR
VAR CONSTANT
    DL_SPP_RMAX : DINT := 32; // 滚动窗容量上界 [拍]，与环形数组一致 / the ring capacity aligned with the array
END_VAR

// 段 0｜复位沿无条件周期刷新（禁入分支，R7）/ segment 0, the unconditional refresh
rtReset(CLK := bReset); // 复位沿 / the reset edge

// 段 1｜首拍初始化与单拍标志预清（R310 / FB32-1 / R256）/ segment 1, the first scan init and the preset
IF NOT _bInit THEN // 首拍一拍 / the first scan
    _bInit := TRUE; // 置首拍标志 / raise the first scan flag
    _bFault := FALSE; // 故障锁存显式清零 / clear the fault latch explicitly
    _bDevFlt := FALSE; // 偏差锁存显式清零 / clear the deviation latch explicitly
    _bDriftFlt := FALSE; // 漂移锁存显式清零 / clear the drift latch explicitly
    _eState := E_DL_SensorPairPhase.eUseA; // 状态显式落 A 源 / place the state to the source A
    _nFill := 0; // 填充计数显式清零（R243 复位清单）/ clear the filled count explicitly
    _nUsePrev := 0; // 窗长快照置 0，使段 2 变更沿必然触发一次全窗清零 / zero the window snapshot so the change edge clears the ring once
    _fRingSum := 0.0; // 环窗和显式清零 / clear the ring sum explicitly
    _nHead := 0; // 写头显式清零 / clear the write head explicitly
END_IF
IF rtReset.Q THEN // 复位沿（作用域：清双侧锁存 + 迁相位 + 清环窗累计量，R311 声明）/ the reset edge with the declared scope
    _bDevFlt := FALSE; // 清偏差锁存（解除路径：复位沿恒可达，R152 自证）/ clear the deviation latch
    _bDriftFlt := FALSE; // 清漂移锁存 / clear the drift latch
    _eState := E_DL_SensorPairPhase.eUseA; // 迁回 A 源 / back to the source A
    _nFill := 0; // 填充计数清零（R243 复位清单）/ clear the filled count
    _nUsePrev := 0; // 窗长快照置 0 触发一次全窗清零 / zero the window snapshot to force a ring clear
    _fRingSum := 0.0; // 环窗和清零 / clear the ring sum
    _nHead := 0; // 写头清零 / clear the write head
END_IF
_bSw := FALSE; // 切换单拍预清零 / preset the switch bit false
_bWinBad := FALSE; // 钳位标记预清零 / preset the clamp flag false

// 段 2｜非有限闸与窗长钳位（R272 全量点名，边界三二）/ segment 2, the finiteness gate and the window clamp
_bFinA := (fA = fA) AND ((fA - fA) = (fA - fA)); // A 源自反 + 差值判 / the A source tests
_bFinB := (fB = fB) AND ((fB - fB) = (fB - fB)); // B 源自反 + 差值判 / the B source tests
_bFin := _bFinA AND _bFinB
AND (fDevWin = fDevWin) AND ((fDevWin - fDevWin) = (fDevWin - fDevWin))
AND (fDriftLim = fDriftLim) AND ((fDriftLim - fDriftLim) = (fDriftLim - fDriftLim)); // 阈值引脚同判 / the threshold pins tested the same way
_nUse := nTrendWin; // 窗长接管 / take the window length
IF (_nUse < 1) OR (_nUse > DL_SPP_RMAX) THEN // 窗长越域（边界二）/ the window length out of the domain
    _bWinBad := TRUE; // 置钳位标记 / raise the clamp flag
    IF _nUse < 1 THEN // 下界钳位 / the floor clamp
        _nUse := 1; // 钳到一 / clamp to one
    ELSE // 上界钳位 / the ceiling clamp
        _nUse := DL_SPP_RMAX; // 钳到容量 / clamp to the capacity
    END_IF
END_IF

// 段 2b｜窗长变更沿全窗清零（v1.0.1 修 D4：仅清和与写头不足，减项 _afRing[_nHead] 会把陈旧样本重新注入和）/ segment 2b, the full window clear on a length change
IF _nUse <> _nUsePrev THEN // 窗长变更沿（含首拍 _nUsePrev = 0）/ the window length change edge, including the first scan
    _fRingSum := 0.0; // 环窗和清零 / clear the ring sum
    _nHead := 0; // 写头回零 / reset the write head
    _nFill := 0; // 填充计数回零 / reset the filled count
    FOR _nRingIdx := 0 TO DL_SPP_RMAX - 1 DO // 有界遍历全容量（32 项，无死循环风险）/ the bounded traversal over the full capacity
        _afRing[_nRingIdx] := 0.0; // 环元素逐项清零：减项读到零才不会把旧样本扣回和里 / zero every element so the subtract term reads zero instead of a stale sample
    END_FOR
    _nUsePrev := _nUse; // 快照本拍窗长，防重复清零 / snapshot the length to avoid a repeated clear
END_IF

// 段 3｜偏差与漂移判据（闸覆盖全量入参后执行）/ segment 3, the deviation and the drift criteria
IF _bFinA AND _bFinB THEN // 双源有限才判偏差（双源非有限即整段跳过，_nFill 保持不增）/ the deviation judged on two finite sources, otherwise the whole segment is skipped
    _fDev := ABS(fA - fB); // 偏差（无除法，无除零风险）/ the deviation without a division
    _fRingSum := _fRingSum - _afRing[_nHead] + _fDev; // 环窗和滑窗更新（环元素已在清零沿置零，减项必为有效样本或零）/ update the ring sum, the subtract term is either a live sample or zero
    _afRing[_nHead] := _fDev; // 本拍偏差入环 / push the deviation into the ring
    _nHead := _nHead + 1; // 写头推进 / advance the head
    IF _nHead >= _nUse THEN // 回卷（按钳位窗长）/ wrap by the clamped length
        _nHead := 0; // 写头回零 / reset the head
    END_IF
    IF _nFill < _nUse THEN // 窗未填满才累加 / count only while the window is not yet full
        _nFill := _nFill + 1; // 填充计数推进 / advance the filled count
    END_IF
    IF _fDev > fDevWin THEN // 偏差超窗（0707 独立成因）/ the deviation over the window
        _bDevFlt := TRUE; // 独立锁存 / latch the deviation cause
    END_IF
    // 除子证明（v1.0.1 重写）：① _nFill 在上一行刚自增且上界为 _nUse，而 _nUse 已在段 2 钳到 ≥ 1，
    // 故进入本判时 _nFill ≥ 1 恒成立；② 唯一能把 _nFill 置 0 的是段 2b 的窗长变更沿，它在段 3 之前执行；
    // ③ 下方 _nFill ≥ 1 复检为第三重防御，供后续重构时不破除零。
    // divisor proof: the count is incremented just above and bounded by the clamped length of at least one, so it is at least one here;
    // the only zeroing path is the length change edge executed before this segment; the explicit recheck below is a third line of defence.
    IF _nFill >= 1 THEN // 除零复检（正常路径恒真，禁用裸除子）/ the divisor recheck, always true on the normal path
        IF (_fRingSum / DINT_TO_LREAL(_nFill)) > fDriftLim THEN // 滚动均值超限（除子已证 ≥ 1，0708 独立成因）/ the rolling mean over the limit with a proven divisor
            _bDriftFlt := TRUE; // 独立锁存 / latch the drift cause
        END_IF
    END_IF
END_IF
IF _bDevFlt OR _bDriftFlt THEN // 任一成因锁存即整体故障 / any cause latches the whole fault
    _bFault := TRUE; // 总锁存 / latch the total fault
END_IF

// 段 4｜择优状态机（ENUM + CASE，ELSE 兜底；迟滞纪律，边界一）/ segment 4, the selection machine with the hysteresis
CASE _eState OF
    E_DL_SensorPairPhase.eUseA: // A 源相 / the source A phase
        IF _bFault THEN // 故障迁移（安全相带全量闸位复检，R274）/ the fault migration with the full gate recheck
            _eState := E_DL_SensorPairPhase.eFault; // 迁入故障锁存相 / enter the fault phase
        ELSIF NOT _bFinA THEN // A 源失效：迟滞边界切换（唯一切换判据）/ the A source invalid, the hysteresis boundary switch
            _eState := E_DL_SensorPairPhase.eUseB; // 切到 B 源 / switch to the source B
            _bSw := TRUE; // 置切换单拍 / raise the switch bit
        END_IF
    E_DL_SensorPairPhase.eUseB: // B 源相 / the source B phase
        IF _bFault THEN // 故障迁移 / the fault migration
            _eState := E_DL_SensorPairPhase.eFault; // 迁入故障锁存相 / enter the fault phase
        ELSIF NOT _bFinB THEN // B 源失效：切回 A / the B source invalid, back to A
            _eState := E_DL_SensorPairPhase.eUseA; // 切回 A 源 / back to the source A
            _bSw := TRUE; // 置切换单拍 / raise the switch bit
        END_IF
    E_DL_SensorPairPhase.eFault: // 故障锁存相：等复位沿（解除可达，边界四）/ the fault phase until the reset edge
        IF rtReset.Q AND (NOT _bDevFlt) AND (NOT _bDriftFlt) THEN // 双锁存已清才迁出（防清锁同拍重锁，FB50-1）/ the exit only after both latches cleared
            _eState := E_DL_SensorPairPhase.eUseA; // 迁回 A 源 / back to the source A
        END_IF
    ELSE // 非法枚举值拦截 / the illegal enumeration guard
        _eState := E_DL_SensorPairPhase.eUseA; // 落回 A 源 / force back to A
        _bFault := TRUE; // 置总锁存 / latch the total fault
END_CASE

// 段 5｜统一出口（择优值按态取源；故障冻结快照，R273）/ segment 5, the unified outlet
bSwitched := _bSw; // 切换单拍出口 / the switch pulse outlet
eState := _eState; // 状态出口 / the state outlet
bSrcA := (_eState = E_DL_SensorPairPhase.eUseA); // A 源指示 / the A indicator
bSrcB := (_eState = E_DL_SensorPairPhase.eUseB); // B 源指示 / the B indicator
IF _eState = E_DL_SensorPairPhase.eUseA THEN // A 源相出口取 A（非有限时安全零，R273）/ the A outlet with the safe zero on a non finite source
    IF _bFinA THEN // A 有限才外泄 / export only a finite A
        fSel := fA; // 择优值 / the selected value
        _fSnap := fA; // 快照更新（写前过闸，FB32-7）/ update the snapshot gated
    ELSE // A 非有限：保持快照（切换已在状态机发生）/ keep the snapshot
        fSel := _fSnap; // 冻结快照出口 / freeze the snapshot outlet
    END_IF
ELSIF _eState = E_DL_SensorPairPhase.eUseB THEN // B 源相出口取 B / the B outlet
    IF _bFinB THEN // B 有限才外泄 / export only a finite B
        fSel := fB; // 择优值 / the selected value
        _fSnap := fB; // 快照更新 / update the snapshot
    ELSE // B 非有限：保持快照 / keep the snapshot
        fSel := _fSnap; // 冻结快照出口 / freeze the snapshot outlet
    END_IF
ELSE // 故障相：冻结最近有效快照（R273）/ the fault phase freezes the snapshot
    fSel := _fSnap; // 冻结快照出口 / freeze the snapshot outlet
END_IF
bError := _bFault; // 故障位出口（与锁存同源）/ the fault bit outlet
bValid := (NOT _bFault) AND (_bFinA OR _bFinB); // 可用标志（无故障且至少一源有限，单点单写）/ the usable flag, no fault and at least one finite source
IF _bDevFlt THEN // 偏差成因回放（R187 锁存回放）/ the deviation cause replayed
    eErr := 16#0003_0707; // 故障级：偏差超窗 / fault grade, the deviation over the window
ELSIF _bDriftFlt THEN // 漂移成因 / the drift cause
    eErr := 16#0003_0708; // 故障级：漂移趋势超限 / fault grade, the drift over the limit
ELSIF _bSw THEN // 切换（信息级不置 bError，R285）/ the switch informational
    eErr := 16#0003_0709; // 信息级：发生择优源切换 / informational, the source switched
ELSIF _bWinBad THEN // 窗长钳位（信息级）/ the window clamp informational
    eErr := 16#0003_070A; // 信息级：滚动窗长度越域已钳位 / informational, the window clamped
ELSE // 无事件 / no event
    eErr := 16#0000_0000; // 正常 / ok
END_IF
END_FUNCTION_BLOCK

(* ---- FB_DL_SensorSupplyWatch.st ---- *)
//==============================================================================
// 功能块：FB_DL_SensorSupplyWatch ｜ 中文名称：传感器供电电压窗口监视
// 所属子库：DL_Device ｜ 版本：v1.0.1 ｜ 日期：2026-11-23
// 兼容：CODESYS V3.5+ / TwinCAT 3 / 汇川 InoProShop（纯 IEC 61131-3，零方言）
// 功能描述：传感器供电电压窗口监视：欠压/过压分级判出（越窗经 tDebounce
//           去抖确认才声明；恢复回正常同样需在窗连续 tDebounce，故障/恢复
//           同一去抖口径，R73 返修），出口按 NE43 四态约定（00 = 正常 /
//           01 = 工作但不正常 / 11 = 故障 / 10 = 无诊断）输出枚举与双 BOOL。
//           窗口参数引脚注入（fVMin / fVMax），非魔法数。
//           同族分工：多通道窗口均值 + 迟滞判限（逐通道掩码诊断）属
//           FB_DL_SensorSupplyMon；本件为单通道供电窗口 NE43 四态监视，
//           互不替代（R73 互引）。
// 开源溯源 (Origin)：候选队列 WINDOW2（oscatBasic，MIT 许可，
//           https://github.com/tkucic/brOscatLib/blob/main/oscatBasic/WINDOW2.st）
//           ——窗口比较行为定义参考；原名 WINDOW2 → 道莅
//           FB_DL_SensorSupplyWatch，clean-room 独立重写（去抖确认 + NE43
//           出口为道莅防御规范增量，零源码行复制）
// 公开接口清单：输入 fSupplyV / fVMin / fVMax / tDebounce；
//               输出 bSupplyOk / bUnder / bOver / eN43 / uErrCode / bValid
// 错误码表：16#0003_0750 信息级（输入非有限判无效，NE43 报 11 故障态，
//           不置 bError——供电异常是工况事实非软件故障）/
//           16#0003_0751 预留禁用（不得挪用）
// 状态机：E_DL_N43State（本文件唯一定义，全库唯一属主，NE43 四态口径）：
//           eOk = 0 / eUnderRange = 1 / eOverRange = 2 / eInvalid = 3
// 边界行为：① 输入非有限 → eInvalid（NE43 = 11 故障态）+ 信息码；
//           ② 越窗经 tDebounce 去抖确认才置 bUnder/bOver（抖动不误报）；
//             恢复回正常同样经在窗去抖 tonOk 确认（同口径，R73 返修）；
//           ③ fVMax <= fVMin 参数倒置 → 视配置故障按 eInvalid 处理；
//           ④ TON ×2 每拍无条件刷新（不入分支，红线 R7）；
//           ⑤ CASE 带 ELSE 非法态兜底归 eInvalid。
// 修订历史：v1.0.0 2026-11-23 首版（R73 派单 · 批 3 · 序 15）
//           v1.0.1 2026-11-23 R73 返修：恢复判定并入故障判定同一去抖口径
//           （新增 tonOk 在窗去抖 + bInOk 暂存，bSupplyOk 改由统一出口按
//           eN43 = eOk 声明）；并补与 FB_DL_SensorSupplyMon 的同族分工互引。
//==============================================================================

(*------------------------------------------------------------------------------
 * 枚举: E_DL_N43State（归属本功能块，同文件发布，全库唯一属主）
 * 含义: NE43 四态诊断出口口径，成员与 CASE 标签双向完备。
 *-----------------------------------------------------------------------------*)
TYPE E_DL_N43State :
(
    eOk         := 0,   // NE43 = 00：正常 / Normal
    eUnderRange := 1,   // NE43 = 01：欠压（工作但不正常）/ Undervoltage, working but not normal
    eOverRange  := 2,   // NE43 = 01：过压（工作但不正常）/ Overvoltage, working but not normal
    eInvalid    := 3    // NE43 = 11：无效/故障（输入非有限或参数倒置）/ Invalid or fault
);
END_TYPE

(*==============================================================================
 * 功能块: FB_DL_SensorSupplyWatch
 * 调用约定: 每个扫描周期无条件调用一次；实例状态全部驻留于私有变量。
 *==============================================================================*)
FUNCTION_BLOCK FB_DL_SensorSupplyWatch
VAR_INPUT
    fSupplyV  : LREAL := 24.0;         // 供电电压实测值 [伏特] / Measured supply voltage [V]
    fVMin     : LREAL := 21.6;         // 电压窗口下限 [伏特]，引脚注入 / Voltage window floor [V], injected via the pin
    fVMax     : LREAL := 26.4;         // 电压窗口上限 [伏特]，引脚注入 / Voltage window ceiling [V], injected via the pin
    tDebounce : TIME  := T#500MS;      // 越窗去抖确认延时 [毫秒] / Out-of-window debounce delay [ms]
END_VAR
VAR_OUTPUT
    bSupplyOk : BOOL;                  // 供电正常声明（去抖后）/ Supply normal declaration after debounce
    bUnder    : BOOL;                  // 欠压声明（去抖确认后）/ Undervoltage declared after debounce
    bOver     : BOOL;                  // 过压声明（去抖确认后）/ Overvoltage declared after debounce
    eN43      : E_DL_N43State;         // NE43 四态出口 / NE43 four-state outlet
    uErrCode  : UDINT;                 // 信息级码，0 = 无信息 / Info-level code, 0 = none
    bValid    : BOOL;                  // 输出可用标志 / Outputs usable flag
END_VAR
VAR
    tonUnder  : TON;                   // 欠压去抖定时器，每拍无条件刷新 / Undervoltage debounce timer, refreshed every scan
    tonOver   : TON;                   // 过压去抖定时器，每拍无条件刷新 / Overvoltage debounce timer, refreshed every scan
    tonOk     : TON;                   // 在窗恢复去抖定时器，每拍无条件刷新 / In-window recovery debounce timer, refreshed every scan
    bInUnder  : BOOL;                  // 本拍欠压越窗（未确认）/ Undervoltage window violation this scan, unconfirmed
    bInOver   : BOOL;                  // 本拍过压越窗（未确认）/ Overvoltage window violation this scan, unconfirmed
    bInOk     : BOOL;                  // 本拍在窗暂存（恢复去抖输入）/ In-window staged this scan, recovery debounce input
    bParamBad : BOOL;                  // 参数倒置声明 / Parameter inversion flag
END_VAR
VAR CONSTANT
    DL_SSV_INF   : LREAL := 1.7976931348623157E308; // LREAL 幅值上限 / LREAL magnitude ceiling
    DL_SSV_CODE_INV : UDINT := 16#0003_0750; // 信息级：输入非有限或参数倒置码 / Info code: non-finite input or inverted parameters
END_VAR

// ---- 段 1｜定时器无条件刷新（红线 R7：禁入条件分支）----
tonUnder(IN := bInUnder, PT := tDebounce); // 欠压去抖按越窗态断输入 / Under timer input per violation state
tonOver(IN := bInOver, PT := tDebounce);   // 过压去抖按越窗态断输入 / Over timer input per violation state
tonOk(IN := bInOk, PT := tDebounce);       // 在窗恢复去抖按在窗态断输入 / Ok timer input per in-window state

// ---- 段 2｜出口默认值：入口即赋确定值 ----
bSupplyOk := FALSE;                   // 正常声明默认 FALSE / Normal declaration preset FALSE
bUnder    := FALSE;                   // 欠压声明默认 FALSE / Undervoltage preset FALSE
bOver     := FALSE;                   // 过压声明默认 FALSE / Overvoltage preset FALSE
bInUnder  := FALSE;                   // 越窗暂存先清零 / Violation stage cleared first
bInOver   := FALSE;                   // 越窗暂存先清零 / Violation stage cleared first
bInOk     := FALSE;                   // 在窗暂存先清零 / In-window stage cleared first
bParamBad := FALSE;                   // 参数倒置声明先清零 / Parameter inversion preset FALSE
uErrCode  := 16#0000_0000;            // 信息码每拍重算（信息级不锁存）/ Info code recomputed, never latched
bValid    := TRUE;                    // 可用标志默认 TRUE / Usable flag preset TRUE
// 注：eN43 为跨拍状态量，不在此预置（初始值 = eOk，由段 5 状态机推进）
// Note: eN43 is a cross-scan state, preset skipped here, advanced by the segment-5 machine

// ---- 段 3｜输入防御与参数闸：非有限或窗口倒置 → eInvalid（NE43 = 11）----
IF (fSupplyV <> fSupplyV) OR (ABS(fSupplyV) > DL_SSV_INF)
   OR (fVMin <> fVMin) OR (ABS(fVMin) > DL_SSV_INF)
   OR (fVMax <> fVMax) OR (ABS(fVMax) > DL_SSV_INF)
   OR (fVMax <= fVMin) THEN
    bParamBad := (fVMax <= fVMin) OR (fVMin <> fVMin) OR (fVMax <> fVMax); // 参数倒置归因 / Parameter inversion attribution
    eN43     := E_DL_N43State.eInvalid; // NE43 故障态 / NE43 invalid state
    uErrCode := DL_SSV_CODE_INV;        // 信息级留痕（不置 bError）/ Info trace, no fault flag
    bValid   := TRUE;                   // 出口确定（无效是合法诊断结论）/ Outlets deterministic
    RETURN;                             // 结构早退（去抖声明保持 FALSE）/ early exit
END_IF

// ---- 段 4｜窗口比较（WINDOW2 行为定义口径）：越窗暂存，去抖确认 ----
IF fSupplyV < fVMin THEN
    bInUnder := TRUE;                   // 欠压越窗暂存 / Undervoltage violation staged
ELSIF fSupplyV > fVMax THEN
    bInOver := TRUE;                    // 过压越窗暂存 / Overvoltage violation staged
END_IF
bUnder    := tonUnder.Q;               // 欠压去抖确认声明 / Undervoltage confirmed
bOver     := tonOver.Q;               // 过压去抖确认声明 / Overvoltage confirmed
bInOk     := (NOT bInUnder) AND (NOT bInOver); // 本拍在窗暂存（恢复去抖输入）/ In-window staged, recovery debounce input

// ---- 段 5｜NE43 出口装配（CASE 带 ELSE；非法态兜底归 eInvalid）----
CASE eN43 OF
    E_DL_N43State.eOk:                 // 正常相：双向未确认越窗
        IF bUnder THEN
            eN43 := E_DL_N43State.eUnderRange; // 升欠压态 / Rise to undervoltage
        ELSIF bOver THEN
            eN43 := E_DL_N43State.eOverRange;  // 升过压态 / Rise to overvoltage
        END_IF
    E_DL_N43State.eUnderRange:         // 欠压态：可升过压或经在窗去抖回正常
        IF bOver THEN
            eN43 := E_DL_N43State.eOverRange;  // 升过压态 / Rise to overvoltage
        ELSIF tonOk.Q THEN                 // 恢复闸：在窗连续 tDebounce 才回正常（与故障判定同口径，R73）/ Recovery gate, same debounce discipline
            eN43 := E_DL_N43State.eOk;         // 回正常态 / Back to normal
        END_IF
    E_DL_N43State.eOverRange:          // 过压态：可落欠压或经在窗去抖回正常
        IF bUnder THEN
            eN43 := E_DL_N43State.eUnderRange; // 落欠压态 / Fall to undervoltage
        ELSIF tonOk.Q THEN                 // 恢复闸：同口径（R73）/ Recovery gate, same discipline
            eN43 := E_DL_N43State.eOk;         // 回正常态 / Back to normal
        END_IF
    E_DL_N43State.eInvalid:            // 无效态：输入恢复合法后按同口径去抖迁移（段 3 早退承担整拍重评）
        IF bUnder THEN
            eN43 := E_DL_N43State.eUnderRange; // 恢复欠压态（去抖确认后）/ Recover to undervoltage after debounce
        ELSIF bOver THEN
            eN43 := E_DL_N43State.eOverRange;  // 恢复过压态（去抖确认后）/ Recover to overvoltage after debounce
        ELSIF tonOk.Q THEN                     // 恢复闸：在窗连续 tDebounce（同口径，R73）/ Recovery gate, same discipline
            eN43 := E_DL_N43State.eOk;         // 恢复正常态 / Recover to normal
        END_IF                                 // 未满任一确认窗：滞留 eInvalid / Stay invalid until a window completes
    ELSE                               // 非法态兜底（R21：CASE 必带 ELSE）
        eN43 := E_DL_N43State.eInvalid; // 拦截非法值归无效态 / Catch illegal value to invalid
END_CASE

// ---- 段 6｜统一出口：正常声明按 NE43 态装配（恢复经 tonOk 去抖后才成立，R73）----
bSupplyOk := (eN43 = E_DL_N43State.eOk); // 正常 = 仅 NE43 正常态（双向去抖同口径）/ Normal = NE43 ok state only, both directions debounced
END_FUNCTION_BLOCK

(* ---- FB_DL_ShearBladeGapSeq.st ---- *)
(*
  Name: FB_DL_ShearBladeGapSeq
  Category: DL_Device
  Version: 1.0.0
  Round: R89 / 2026-11-25
  开源溯源：clean-room 自研（族 板带剪切分条卷取，ST 开源生态实测 0 命中，无外部代码引入）
  功能：剪切刀间隙调整与锁定顺控：松开夹紧→伺服调隙→间隙测量确认→夹紧锁定。
  边界条件：① 位置与公差入参全部过非有限闸；配置越域即故障（101）；
            ② 松开/调整/确认/夹紧四相各用独立 TON，PT 均取 tTimeoutS，禁跨相共用（R100）；
            ③ 确认相要求「偏差在带内且仍处于松开状态」，防夹紧前已被误夹导致间隙失真；
            ④ 故障解除唯一路径：故障相内 xStart 释放（R152），清锁存回 eIdle。
  状态机：eIdle / eRelease / eAdjust / eVerify / eClamp / eDone / eFault（CASE 含 ELSE 兜底）。
*)
TYPE E_DL_SbgPhase :
(
    eIdle    := 0,      (* 待机：等启动沿 / Idle, waiting for start edge *)
    eRelease := 10,     (* 松开相：等夹紧松开反馈 / Release, waiting clamp open *)
    eAdjust  := 20,     (* 调整相：伺服调隙进带 / Adjusting gap into band *)
    eVerify  := 30,     (* 确认相：测量确认且仍松开 / Verify gap while still released *)
    eClamp   := 40,     (* 夹紧相：等夹紧到位 / Clamping, waiting lock feedback *)
    eDone    := 50,     (* 完成相：保持至启动释放 / Done, holds until start released *)
    eFault   := 90      (* 故障相：锁存待释放 / Fault latched, awaiting release *)
);
END_TYPE

FUNCTION_BLOCK FB_DL_ShearBladeGapSeq
VAR_INPUT
    xStart : BOOL;          (* 启动命令（上升沿起序） [-] Start command, rising edge *)
    fGapTargetMm : REAL;    (* 间隙目标值 [mm] Target gap [mm] *)
    fGapActMm : REAL;       (* 间隙实测值 [mm] Actual gap [mm] *)
    fGapTolMm : REAL;       (* 间隙公差 [mm] Gap tolerance [mm] *)
    xClamped : BOOL;        (* 夹紧到位反馈（TRUE = 已夹紧） [-] Clamp feedback *)
    tTimeoutS : TIME;       (* 单相超时窗 [ms] Phase timeout window [ms] *)
END_VAR
VAR_OUTPUT
    eState : E_DL_SbgPhase; (* 当前相 [-] Present phase *)
    xDone : BOOL;           (* 完成单拍脉冲 [-] One-scan done pulse *)
    xFault : BOOL;          (* 故障锁存标志 [-] Fault latched *)
    nErrCode : INT;         (* 故障码 0/101 组态/102~105 超时/106 非法相 [-] Error code *)
END_VAR
VAR
    _ePhase : E_DL_SbgPhase := E_DL_SbgPhase.eIdle;  (* 内部相（CASE 唯一写入目标） [-] Internal phase *)
    _bDone : BOOL := FALSE;         (* 单拍完成标志（段 1 预清） [-] One-scan done flag *)
    _bFaultLatch : BOOL := FALSE;   (* 故障锁存位 [-] Fault latch *)
    _bReqFault : BOOL := FALSE;     (* 单拍故障请求（段 1 预清） [-] Fault request *)
    _bCfgBad : BOOL := FALSE;       (* 组态非法当拍量 [-] Configuration bad *)
    _nErr : INT := 0;               (* 故障码锁存 [-] Latched error code *)
    _nReqErr : INT := 0;            (* 当拍请求码 [-] Requested error code *)
    _fErrMm : REAL := 0.0;          (* 间隙偏差绝对量 [mm] Absolute gap deviation [mm] *)
    tonRelease : TON;               (* 松开超时（段 0 无条件调用） / Release timeout *)
    tonAdjust : TON;                (* 调整超时（段 0 无条件调用） / Adjust timeout *)
    tonVerify : TON;                (* 确认超时（段 0 无条件调用） / Verify timeout *)
    tonClamp : TON;                 (* 夹紧超时（段 0 无条件调用） / Clamp timeout *)
    rtStart : R_TRIG;               (* 启动沿（段 0 无条件调用） / Start edge *)
END_VAR
VAR CONSTANT
    DL_SBG_EPS : REAL := 1.0E-9;    (* 判据容差 [-] Criterion tolerance *)
END_VAR
(* —— 段 0：沿与四 TON 无条件周期刷新（R7），IN 仅由相位派生 —— *)
rtStart(CLK := xStart);                                                     (* 启动沿 / Start edge *)
tonRelease(IN := (_ePhase = E_DL_SbgPhase.eRelease), PT := tTimeoutS);      (* 松开超时 / Release timeout *)
tonAdjust(IN := (_ePhase = E_DL_SbgPhase.eAdjust), PT := tTimeoutS);        (* 调整超时 / Adjust timeout *)
tonVerify(IN := (_ePhase = E_DL_SbgPhase.eVerify), PT := tTimeoutS);        (* 确认超时 / Verify timeout *)
tonClamp(IN := (_ePhase = E_DL_SbgPhase.eClamp), PT := tTimeoutS);          (* 夹紧超时 / Clamp timeout *)
(* 非有限闸（NaN 自反 + Inf 差值自减）+ 组态域闸：三浮点入参全枚举（R272） *)
_bCfgBad := (fGapTargetMm <> fGapTargetMm) OR ((fGapTargetMm - fGapTargetMm) <> 0.0)
         OR (fGapActMm <> fGapActMm) OR ((fGapActMm - fGapActMm) <> 0.0)
         OR (fGapTolMm <> fGapTolMm) OR ((fGapTolMm - fGapTolMm) <> 0.0)
         OR (fGapTargetMm <= 0.0) OR (fGapTargetMm > 50.0)
         OR (fGapTolMm <= DL_SBG_EPS) OR (fGapTolMm > 5.0) OR (tTimeoutS <= T#0S);
(* 偏差绝对量：容差比较一律用差值，禁浮点判等 *)
_fErrMm := ABS(fGapActMm - fGapTargetMm);
(* —— 段 1：单拍量预清零 —— *)
_bDone := FALSE;
_bReqFault := FALSE;
_nReqErr := 0;
IF _bCfgBad THEN
    _bReqFault := TRUE; _nReqErr := 101;        (* 组态非法 / Configuration bad *)
END_IF
(* —— 段 2：故障锁存解除（唯一路径 = 故障相内 xStart 释放，R152） —— *)
IF _bFaultLatch AND (NOT xStart) THEN
    _bFaultLatch := FALSE;                      (* 清锁存 / Clear latch *)
    _nErr := 0;                                 (* 清码 / Clear code *)
    _ePhase := E_DL_SbgPhase.eIdle;             (* 迁回待机 / Back to idle *)
END_IF
(* —— 段 3：主状态机（ENUM + CASE，ELSE 兜底） —— *)
CASE _ePhase OF
E_DL_SbgPhase.eIdle:
    IF rtStart.Q AND (NOT _bFaultLatch) THEN
        _ePhase := E_DL_SbgPhase.eRelease;      (* 起序 → 松开 / Start to release *)
    END_IF
E_DL_SbgPhase.eRelease:
    IF NOT xClamped THEN
        _ePhase := E_DL_SbgPhase.eAdjust;       (* 已松开 → 调隙 / Released, adjust *)
    ELSIF tonRelease.Q THEN
        _bReqFault := TRUE; _nReqErr := 102;    (* 松开超时 / Release timeout *)
    END_IF
E_DL_SbgPhase.eAdjust:
    IF _fErrMm <= fGapTolMm THEN
        _ePhase := E_DL_SbgPhase.eVerify;       (* 进带 → 测量确认 / In band, verify *)
    ELSIF tonAdjust.Q THEN
        _bReqFault := TRUE; _nReqErr := 103;    (* 调整超时 / Adjust timeout *)
    END_IF
E_DL_SbgPhase.eVerify:
    IF (_fErrMm <= fGapTolMm) AND (NOT xClamped) THEN
        _ePhase := E_DL_SbgPhase.eClamp;        (* 确认通过且仍松开 → 夹紧 / Verified, clamp *)
    ELSIF tonVerify.Q THEN
        _bReqFault := TRUE; _nReqErr := 104;    (* 确认超时 / Verify timeout *)
    END_IF
E_DL_SbgPhase.eClamp:
    IF xClamped AND (_fErrMm <= fGapTolMm) THEN
        _bDone := TRUE;                         (* 单拍完成（段 1 预清） / One-scan done *)
        _ePhase := E_DL_SbgPhase.eDone;         (* → 完成相 / To done *)
    ELSIF tonClamp.Q THEN
        _bReqFault := TRUE; _nReqErr := 105;    (* 夹紧超时 / Clamp timeout *)
    END_IF
E_DL_SbgPhase.eDone:
    IF NOT xStart THEN
        _ePhase := E_DL_SbgPhase.eIdle;         (* 启动释放 → 待机 / Start released, idle *)
    END_IF
E_DL_SbgPhase.eFault:
    _fErrMm := ABS(fGapActMm - fGapTargetMm);   (* 故障相驻留：仅刷新偏差量供追溯，不迁相 *)
ELSE
    _bReqFault := TRUE;                         (* 非法相兜底 / Illegal phase fallback *)
    _nReqErr := 106;
END_CASE
(* —— 段 4：故障请求统一落地（唯一锁存点 + 同步迁相，R187/R252） —— *)
IF _bReqFault AND (NOT _bFaultLatch) THEN
    _bFaultLatch := TRUE;                       (* 锁存 / Latch *)
    _nErr := _nReqErr;                          (* 码锁存回放 / Latched code *)
    _ePhase := E_DL_SbgPhase.eFault;            (* 同步迁相 / Migrate to fault *)
END_IF
(* —— 段 5：统一出口（各出口单点赋值） —— *)
eState := _ePhase;
xDone := _bDone;
xFault := _bFaultLatch;
nErrCode := _nErr;
END_FUNCTION_BLOCK

(* ---- FB_DL_SingleSolenoidCyl.st ---- *)
(*==============================================================================
 * 组件名称 (Component)  : FB_DL_SingleSolenoidCyl
 * 所属子库 (Sublibrary) : DL_Device
 * 当前版本 (Version)    : 1.0.1
 * 兼容性   (Platform)   : CODESYS 3.5 / TwinCAT 3 / 汇川 InoProShop / Machine Expert
 *                         仅依赖 Standard.library（TON / R_TRIG）与 DL_Base
 *                         的 FB_DL_SignalDebounce，零厂商方言
 * 分类     (Category)   : 设备执行器功能块（Function Block，实现 I_DL_Cylinder）
 * 功能简述 (Function)   : 单电控（单线圈）弹簧复位气缸驱动。得电伸出、失电
 *                         弹簧缩回；无传感器纯时间模式 + 可选磁开关反馈
 *                         双重校验模式；联锁中途撤除线圈失电弹簧复位；
 *                         出口断言保证故障/空闲稳态线圈必断；行程计数；
 *                         状态机复用既有 E_DL_CylinderState（禁止重定义），
 *                         ENUM + CASE + ELSE 兜底。
 * 接口实现 (Implements) : I_DL_Cylinder。接口 OUT 列同名成员（eState/
 *                         bExtended/bRetracted/bFault/uErrorId）按 R22 以
 *                         只读 PROPERTY GET 承载（内部镜像同源，非接口
 *                         成员 bSolenoidExt/bMoving/uCycleCount 保留
 *                         VAR_OUTPUT）；方法 CmdExtend/CmdRetract/CmdStop/
 *                         CmdReset 全部在本文件尾部落地。
 * 开源溯源 (Origin)     : 来源标签 lbp-device（RAW_NOTES_R6 S-1：单电控弹簧
 *                         复位气缸的纯时间定位 + 磁开校验双模式、单线圈
 *                         失电即缩回的保位语义等行业公知工程惯例，公开教学
 *                         资料，仅借鉴通用工程语义；状态机、故障码按本库
 *                         红线独立设计，clean-room 未复制源码）。
 * 红线自检 (Redline)    : R1 零全局变量表/外部变量引用 ✓｜R2 零物理 IO 地址 ✓
 *                         R3 纯 IEC 61131-3 ✓｜R4 防越界/出口断言 ✓
 *                         R5 全变量中英双语同行注释 ✓｜R6 ENUM+CASE+ELSE ✓
 *                         R7 九个定时器/边缘/消抖实例主体最前部无条件刷新 ✓
 * 公约遵循 (Convention) : 0.1/R23 本块为纯事件型状态机（BOOL 指令/反馈 +
 *                         TIME 参数，无积分/滤波类连续量同步语义），免首扫，
 *                         无内部初始化标志。
 *                         0.7 故障码段位 16#0003_xxxx：【故障级】0003_0220
 *                         伸出到位超时 / 0003_0221 反馈校验失败 / 0003_0222
 *                         非法状态，全部 R15 锁存仅复位可清；本块无信息级
 *                         码，bFault 派生式天然排除信息级（0.2）。
 * 偏离留档 (Deviation)  : 依 R11 头注释留档，共 2 条：
 *                         ① 规格中 0003_0221 释义"时间到位但磁开超窗未确认"
 *                           与 0003_0220（伸出到位超时）在伸出方向同窗重叠；
 *                           本实现将 0221 明确用于缩回方向的磁开校验超窗
 *                           （弹簧复位时间到位后磁开仍未确认），两码位各自
 *                           可测、语义不冲突。
 *                         ② bCmdExtend 规格标注"上升沿生效"，因单线圈物理
 *                           语义为"得电即伸出、失电即缩回"（电平跟随），
 *                           本实现按 电平 OR 上升沿 双通道受理，电平语义
 *                           自然涵盖边沿语义，不会产生指令保持而线圈断开
 *                           的悬挂态。
 * 修订历史 (Revision)   :
 *   2026-11-15  v1.0.0  首版入库（R6 轮 · DL_Device 阀门/驱动族深化）
 *   2026-11-15  v1.0.1  R11 修复：变量名勘误，段 2 行程计数赋值目标
 *                       _uCycleCount → uCycleCount（原写下划线前缀但未在
 *                       VAR 区声明，且同名输出 uCycleCount 全文零写入，
 *                       判定为前缀笔误而非缺声明；三平台编译阻断已消除）。
 *                       R11 fix: name erratum, _uCycleCount -> uCycleCount
 *============================================================================*)
FUNCTION_BLOCK FB_DL_SingleSolenoidCyl IMPLEMENTS I_DL_Cylinder
VAR_INPUT
    bCmdExtend      : BOOL;           // 伸出指令（Extend command），电平 OR 上升沿双通道受理；失电即弹簧缩回 / Extend command, level or edge accepted, coil drop means spring return
    bSnsExtended    : BOOL;           // 可选伸出到位磁性开关（Optional extended reed switch），TRUE=到位；未接时恒 FALSE / Optional extended reed switch, TRUE = in position, FALSE if not wired
    bSnsRetracted   : BOOL;           // 可选缩回到位磁性开关（Optional retracted reed switch），TRUE=到位 / Optional retracted reed switch, TRUE = in position
    bUseSensorCheck : BOOL;           // 反馈校验使能（Sensor check enable），TRUE=时间+磁开双重校验；FALSE=纯时间模式 / Sensor check enable, TRUE = time + reed dual check, FALSE = pure time mode
    bInterlock      : BOOL;           // 允许动作联锁（Motion interlock），TRUE=允许伸出，默认 FALSE 线圈保持断开 / Motion interlock, TRUE = extend allowed, default FALSE holds coil off
    tStrokeTimeExt  : TIME := T#1S;   // 伸出行程时间（Extend stroke time），纯时间模式据此判定到位 / Extend stroke time, basis of position judgment in pure time mode
    tStrokeTimeRet  : TIME := T#1S;   // 弹簧缩回行程时间（Spring return stroke time），纯时间模式据此判定到位 / Spring return stroke time, basis in pure time mode
    tTimeoutExt     : TIME := T#3S;   // 伸出到位超时（Extend timeout），双重校验模式下磁开确认窗口，T#0S=禁用自检 / Extend timeout for reed confirmation window in dual-check mode, T#0S disables
    tDebounce       : TIME := T#20MS; // 磁开防抖窗口（Sensor debounce），T#0S=直通 / Reed switch debounce window, T#0S = pass-through
    bReset          : BOOL;           // 故障复位（Fault reset），上升沿生效 / Fault reset, rising edge effective
END_VAR

VAR_OUTPUT
    bSolenoidExt  : BOOL;             // 伸出线圈输出（Extend solenoid coil），得电伸出 / 失电弹簧缩回 / Extend solenoid coil, energized to extend, de-energized for spring return
    bMoving       : BOOL;             // 运动中指示（Moving indicator），伸出或缩回动作中 / Moving indicator, while extending or retracting
    uCycleCount   : UDINT;            // 行程计数（Stroke count），缩回判定沿 +1 / Stroke count, incremented on retracted-state edge
END_VAR

VAR
    _eState          : E_DL_CylinderState := E_DL_CylinderState.eIdle; // 内部状态机步序（Internal state step），外部经属性只读 / Internal state, read-only via property
    _bFaultLatch     : BOOL;           // 故障锁存标志（Fault latch flag），仅复位清除 / Fault latch flag, cleared only by reset
    _uErrorIdInt     : UDINT;          // 内部故障码寄存（Internal error register），随锁存写入 / Internal error register written on latch
    _bMethExtLatch   : BOOL;           // 方法伸出保持锁存（Method extend hold latch），由 CmdExtend 置位 / Method extend hold latch set by CmdExtend
    _bMethRetLatch   : BOOL;           // 方法缩回保持锁存（Method retract hold latch），由 CmdRetract/CmdStop 置位 / Method retract hold latch set by CmdRetract or CmdStop
    _bPendStop       : BOOL;           // 方法停止请求（Method stop request），由 CmdStop 置位 / Method stop request set by CmdStop
    _bPendReset      : BOOL;           // 方法复位请求（Method reset request），由 CmdReset 置位 / Method reset request set by CmdReset
    _bExtFilt        : BOOL;           // 消抖后伸出磁开（Debounced extended reed）/ Debounced extended reed signal
    _bRetFilt        : BOOL;           // 消抖后缩回磁开（Debounced retracted reed）/ Debounced retracted reed signal
    _bToEn           : BOOL;           // 磁开确认窗口使能（Confirmation window enable），超时参数大于零时有效 / Confirmation window enable, active when timeout above zero
    _bInStrokeExt    : BOOL;           // 伸出态判定中间量（Extending-state test intermediate），喂定时器实例 / Extending-state test intermediate feeding timer instances
    _bInStrokeRet    : BOOL;           // 缩回态判定中间量（Retracting-state test intermediate），喂定时器实例 / Retracting-state test intermediate feeding timer instances
    _bInExtTo        : BOOL;           // 伸出磁开超时窗计时条件（Ext. reed timeout timing condition）/ Timing condition of extend reed timeout window
    _bInRetFbWin     : BOOL;           // 缩回磁开校验窗计时条件（Ret. reed check window condition），行程时间计满后启动 / Retract reed check window condition, starts after stroke time elapsed
    _bInRetractedSt  : BOOL;           // 已缩回态判定中间量（Retracted-state test intermediate），喂计数边缘实例 / Retracted-state test intermediate feeding count edge instance
    _fbDebExt        : FB_DL_SignalDebounce; // 伸出磁开消抖实例（Extended reed debounce），通道一 / Extended reed debounce instance, channel 1
    _fbDebRet        : FB_DL_SignalDebounce; // 缩回磁开消抖实例（Retracted reed debounce），通道二 / Retracted reed debounce instance, channel 2
    _fbTrigExt       : R_TRIG;         // 引脚伸出指令上升沿（Pin extend command edge）/ Pin extend command rising edge
    _fbTrigReset     : R_TRIG;         // 引脚复位上升沿（Pin reset edge）/ Pin reset rising edge
    _fbTrigRetState  : R_TRIG;         // 进入已缩回态计数上升沿（Retracted-state count edge）/ Rising edge on entering retracted state for stroke counting
    _fbTonStrokeExt  : TON;            // 伸出行程时间定时器（Extend stroke time timer）/ Extend stroke time timer instance
    _fbTonStrokeRet  : TON;            // 弹簧缩回行程时间定时器（Spring return stroke time timer）/ Spring return stroke time timer instance
    _fbTonExtTo      : TON;            // 伸出磁开确认超时定时器（Extend reed confirmation timeout timer）/ Extend reed confirmation timeout timer instance
    _fbTonRetFb      : TON;            // 缩回磁开校验窗定时器（Retract reed check window timer）/ Retract reed check window timer instance
END_VAR

METHOD CmdExtend : BOOL
VAR_INPUT
END_VAR
IF _bFaultLatch OR (_eState = E_DL_CylinderState.eFault) THEN
    CmdExtend       := FALSE;   // 故障态拒绝（Rejected in fault state）
    _bMethRetLatch  := FALSE;   // 清反向残留锁存（Clear stale reverse latch）
ELSE
    _bMethExtLatch  := TRUE;    // 登记伸出保持锁存（Register extend hold latch）
    _bMethRetLatch  := FALSE;   // 互斥注销缩回锁存（Cancel opposite retract latch）
    CmdExtend       := TRUE;    // 受理成功（Accepted）
END_IF

(*------------------------------------------------------------------------------
 * 方法: CmdRetract —— 缩回指令（单线圈释放线圈，弹簧复位）。故障态拒绝。
 *      Method CmdRetract - release coil for spring return, rejected in fault.
 *------------------------------------------------------------------------------*)
    END_METHOD

METHOD CmdRetract : BOOL
VAR_INPUT
END_VAR
IF _bFaultLatch OR (_eState = E_DL_CylinderState.eFault) THEN
    CmdRetract      := FALSE;   // 故障态拒绝（Rejected in fault state）
    _bMethExtLatch  := FALSE;   // 清反向残留锁存（Clear stale reverse latch）
ELSE
    _bMethRetLatch  := TRUE;    // 登记缩回锁存（Register retract latch）
    _bMethExtLatch  := FALSE;   // 互斥注销伸出锁存（Cancel opposite extend latch）
    CmdRetract      := TRUE;    // 受理成功（Accepted）
END_IF

(*------------------------------------------------------------------------------
 * 方法: CmdStop —— 线圈释放、弹簧复位至缩回位（单线圈安全侧）。
 *      Method CmdStop - release coil, spring returns to retracted (safe side).
 *------------------------------------------------------------------------------*)
    END_METHOD

METHOD CmdStop : BOOL
VAR_INPUT
END_VAR
IF _bFaultLatch OR (_eState = E_DL_CylinderState.eFault) THEN
    CmdStop         := FALSE;   // 故障态拒绝（Rejected in fault state）
ELSE
    _bMethExtLatch  := FALSE;   // 注销伸出锁存（Cancel extend latch）
    _bMethRetLatch  := TRUE;    // 登记缩回锁存，主体状态机消化（Register retract latch, consumed by body）
    _bPendStop      := TRUE;    // 登记停止请求（Register stop request）
    CmdStop         := TRUE;    // 受理成功（Accepted）
END_IF

(*------------------------------------------------------------------------------
 * 方法: CmdReset —— 复位故障，返回是否可复位（存在锁存故障时为 TRUE）。
 *      Method CmdReset - reset fault, returns TRUE only when a latch exists.
 *------------------------------------------------------------------------------*)
    END_METHOD

METHOD CmdReset : BOOL
VAR_INPUT
END_VAR
IF _bFaultLatch OR (_eState = E_DL_CylinderState.eFault) THEN
    _bPendReset     := TRUE;    // 登记复位请求，主体状态机消化（Register reset request, consumed by body）
    CmdReset        := TRUE;    // 可复位（Resettable）
ELSE
    CmdReset        := FALSE;   // 无故障可复位（Nothing to reset）
END_IF

(*------------------------------------------------------------------------------
 * 属性: eState（GET）—— 当前状态机状态只读视图。
 *      Property eState (GET) - read-only view of the current state machine state.
 *------------------------------------------------------------------------------*)
    END_METHOD

// ============================================================================
// 段 1｜定时器与边缘检测实例无条件周期刷新（R7：严禁置于 IF/CASE 分支内）
//      Unconditional per-cycle refresh of all timer and edge instances (R7)
// ============================================================================
_fbDebExt(bRawInput := bSnsExtended, tRiseDelay := tDebounce, tFallDelay := tDebounce, bEnable := TRUE, bReset := FALSE);
_fbDebRet(bRawInput := bSnsRetracted, tRiseDelay := tDebounce, tFallDelay := tDebounce, bEnable := TRUE, bReset := FALSE);
_fbTrigExt(CLK := bCmdExtend);
_fbTrigReset(CLK := bReset);
_bExtFilt := _fbDebExt.bStable;       // 通道一消抖输出（Channel 1 debounced output）
_bRetFilt := _fbDebRet.bStable;       // 通道二消抖输出（Channel 2 debounced output）
_bInRetractedSt := (_eState = E_DL_CylinderState.eRetracted); // 已缩回态判定（Retracted-state test）
_fbTrigRetState(CLK := _bInRetractedSt);
_bToEn := (tTimeoutExt > T#0S);       // 窗口参数为零 = 自检禁用（Zero window = check disabled）
_bInStrokeExt := (_eState = E_DL_CylinderState.eExtending);   // 伸出态判定（Extending-state test）
_bInStrokeRet := (_eState = E_DL_CylinderState.eRetracting);  // 缩回态判定（Retracting-state test）
_bInExtTo := _bInStrokeExt AND bUseSensorCheck;               // 双重校验模式才计时确认窗（Window timed only in dual-check mode）
_bInRetFbWin := _bInStrokeRet AND bUseSensorCheck AND _fbTonStrokeRet.Q; // 行程时间计满后启动校验窗（Window starts after stroke time elapsed）
_fbTonStrokeExt(IN := _bInStrokeExt, PT := tStrokeTimeExt);
_fbTonStrokeRet(IN := _bInStrokeRet, PT := tStrokeTimeRet);
_fbTonExtTo(IN := _bInExtTo, PT := tTimeoutExt);
_fbTonRetFb(IN := _bInRetFbWin, PT := tTimeoutExt);

// ============================================================================
// 段 2｜行程计数：进入已缩回态上升沿 +1（纯时间模式同样有效，R15 范畴外）
//      Stroke counting: one increment per retracted-state edge, valid in
//      pure time mode too (outside fault-latch scope)
// ============================================================================
IF _fbTrigRetState.Q THEN
    uCycleCount := uCycleCount + 1; // 完整行程 +1（One completed stroke added）
END_IF

// ============================================================================
// 段 3｜核心状态机（ENUM + CASE，含 ELSE 非法状态兜底）
//      Core state machine (ENUM + CASE with ELSE illegal-state fallback)
// ============================================================================
CASE _eState OF

    E_DL_CylinderState.eIdle: // 空闲稳态：线圈必断，按磁开同步实际位置
        IF _bExtFilt AND (NOT _bRetFilt) THEN
            _eState := E_DL_CylinderState.eExtended;   // 首态同步：实际已伸出（Sync: physically extended）
        ELSIF _bRetFilt AND (NOT _bExtFilt) THEN
            _eState := E_DL_CylinderState.eRetracted;  // 首态同步：实际已缩回（Sync: physically retracted）
        ELSIF (bCmdExtend OR _fbTrigExt.Q OR _bMethExtLatch) AND bInterlock AND (NOT _bMethRetLatch) THEN
            _eState := E_DL_CylinderState.eExtending;  // 受理伸出（Accept extend）
        ELSIF _bMethRetLatch OR _bPendStop THEN
            _bMethRetLatch := FALSE;                   // 空闲态消化缩回/停止请求（Absorb retract/stop requests in idle）
            _bPendStop     := FALSE;
        END_IF

    E_DL_CylinderState.eExtending: // 伸出动作中：线圈得电
        IF bUseSensorCheck AND _bExtFilt AND (NOT _bRetFilt) THEN
            _eState := E_DL_CylinderState.eExtended;   // 双重校验：磁开确认到位（Dual check: reed confirms position）
        ELSIF (NOT bUseSensorCheck) AND _fbTonStrokeExt.Q THEN
            _eState := E_DL_CylinderState.eExtended;   // 纯时间模式：行程时间计满判定到位（Pure time: stroke time elapsed）
        ELSIF bUseSensorCheck AND _bToEn AND _fbTonExtTo.Q THEN
            _bFaultLatch := TRUE;                      // 超时故障锁存（Timeout fault latch）
            _uErrorIdInt := 16#0003_0220;              // 0003_0220 伸出到位超时（磁开窗内未确认）【故障级】/ Extend timeout, fault level
            _eState      := E_DL_CylinderState.eFault;
        ELSIF (NOT (bCmdExtend OR _bMethExtLatch)) OR (NOT bInterlock) THEN
            _eState := E_DL_CylinderState.eRetracting; // 指令失电或联锁中途撤除：线圈断、弹簧复位（Command dropped or interlock removed: coil off, spring return）
        ELSIF _bPendStop OR _bMethRetLatch THEN
            _bPendStop     := FALSE;                   // 停止/缩回请求：线圈断弹簧复位（Stop/retract request: coil off, spring return）
            _bMethExtLatch := FALSE;
            _eState        := E_DL_CylinderState.eRetracting;
        END_IF

    E_DL_CylinderState.eExtended: // 已伸出到位稳态：线圈保持得电维持伸出位
        IF (NOT (bCmdExtend OR _bMethExtLatch)) OR (NOT bInterlock) THEN
            _eState := E_DL_CylinderState.eRetracting; // 指令失电或联锁撤除：失电弹簧缩回（Command dropped or interlock removed: spring return）
        ELSIF _bPendStop OR _bMethRetLatch THEN
            _bPendStop     := FALSE;                   // 停止/缩回请求：失电缩回（Stop/retract request: spring return）
            _bMethExtLatch := FALSE;
            _eState        := E_DL_CylinderState.eRetracting;
        END_IF

    E_DL_CylinderState.eRetracting: // 缩回动作中：线圈失电，弹簧复位不可中断
        IF (NOT bUseSensorCheck) AND _fbTonStrokeRet.Q THEN
            _eState := E_DL_CylinderState.eRetracted;  // 纯时间模式：缩回时间计满（Pure time: return stroke time elapsed）
        ELSIF bUseSensorCheck AND _bRetFilt AND (NOT _bExtFilt) THEN
            _eState := E_DL_CylinderState.eRetracted;  // 双重校验：磁开确认到位（Dual check: reed confirms position）
        ELSIF bUseSensorCheck AND _bToEn AND _fbTonRetFb.Q THEN
            _bFaultLatch := TRUE;                      // 反馈校验失败锁存（Feedback check failure latch）
            _uErrorIdInt := 16#0003_0221;              // 0003_0221 反馈校验失败（缩回时间到位但磁开超窗未确认）【故障级】/ Feedback check failure, fault level
            _eState      := E_DL_CylinderState.eFault;
        ELSIF (bCmdExtend OR _bMethExtLatch) AND bInterlock AND (NOT _bMethRetLatch) THEN
            _eState := E_DL_CylinderState.eExtending;  // 缩回途中再伸出（Re-extend during spring return）
        ELSIF _bPendStop THEN
            _bPendStop := FALSE;                       // 消化停止请求，继续缩回至到位（Absorb stop request, spring return continues）
        END_IF

    E_DL_CylinderState.eRetracted: // 已缩回到位稳态：弹簧保持，线圈必断
        IF _bMethRetLatch THEN
            _bMethRetLatch := FALSE;                   // 缩回锁存到位即消化（Retract latch absorbed at retracted position）
        END_IF
        IF (bCmdExtend OR _fbTrigExt.Q OR _bMethExtLatch) AND bInterlock THEN
            _eState := E_DL_CylinderState.eExtending;  // 受理伸出（Accept extend）
        END_IF

    E_DL_CylinderState.eFault: // 故障锁存态：清空全部请求，仅复位可退出
        _bMethExtLatch := FALSE;                       // 清方法锁存（Clear method latches）
        _bMethRetLatch := FALSE;
        _bPendStop     := FALSE;
        IF _bPendReset OR _fbTrigReset.Q THEN
            _bPendReset  := FALSE;                     // 消费复位请求（Consume reset request）
            _bFaultLatch := FALSE;                     // 解除锁存（Release latch）
            _uErrorIdInt := 0;                         // 故障码清零（Error code cleared）
            _eState      := E_DL_CylinderState.eIdle;  // 回空闲态重新同步（Back to idle for re-sync）
        END_IF

    ELSE // 非法状态兜底：任何越界枚举值强制锁存故障（Illegal state fallback）
        _bFaultLatch := TRUE;                          // 故障锁存（Fault latched）
        _uErrorIdInt := 16#0003_0222;                  // 0003_0222 非法状态【故障级】/ Illegal state, fault level
        _eState      := E_DL_CylinderState.eFault;
END_CASE

// ============================================================================
// 段 4｜线圈输出推导 + 出口断言（硬约束：故障/空闲稳态线圈必断）
//      Coil output derivation + exit assertion (fault/idle states force coil off)
// ============================================================================
bSolenoidExt := (_eState = E_DL_CylinderState.eExtending) OR (_eState = E_DL_CylinderState.eExtended); // 伸出与保持位得电（Energized in extending and extended hold）
IF (_eState = E_DL_CylinderState.eFault) OR (_eState = E_DL_CylinderState.eIdle) THEN
    bSolenoidExt := FALSE;                             // 出口断言：故障/空闲稳态线圈必断（Assertion: coil forced off in fault/idle）
END_IF
bMoving := (_eState = E_DL_CylinderState.eExtending) OR (_eState = E_DL_CylinderState.eRetracting); // 运动中派生（Moving derived）

(*------------------------------------------------------------------------------
 * 方法: CmdExtend —— 伸出指令（登记保持锁存）。故障态一律拒绝返回 FALSE。
 *      Method CmdExtend - register extend hold latch, rejected with FALSE in fault.
 *------------------------------------------------------------------------------*)

PROPERTY eState : E_DL_CylinderState
eState := _eState;            // 返回内部状态（Return internal state）

(*------------------------------------------------------------------------------
 * 属性: bExtended（GET）—— 伸出到位磁开反馈（消抖后）。
 *      Property bExtended (GET) - debounced extended reed feedback.
 *------------------------------------------------------------------------------*)
PROPERTY bExtended : BOOL
bExtended := _bExtFilt;       // 返回通道一消抖输出（Return channel 1 debounced output）

(*------------------------------------------------------------------------------
 * 属性: bRetracted（GET）—— 缩回到位磁开反馈（消抖后）。
 *      Property bRetracted (GET) - debounced retracted reed feedback.
 *------------------------------------------------------------------------------*)
PROPERTY bRetracted : BOOL
bRetracted := _bRetFilt;      // 返回通道二消抖输出（Return channel 2 debounced output）

(*------------------------------------------------------------------------------
 * 属性: bFault（GET）—— 故障锁存指示（信息级码不置本位，0.2 公约）。
 *      Property bFault (GET) - fault latch indicator, info-level codes excluded.
 *------------------------------------------------------------------------------*)
PROPERTY bFault : BOOL
bFault := _bFaultLatch OR (_eState = E_DL_CylinderState.eFault); // 显式排除信息级派生式（Explicit derived form excluding info codes）

(*------------------------------------------------------------------------------
 * 属性: uErrorId（GET）—— 末次故障码（0=无故障）。
 *      Property uErrorId (GET) - last error code (0 = none).
 *------------------------------------------------------------------------------*)
PROPERTY uErrorId : UDINT
uErrorId := _uErrorIdInt;     // 返回内部故障码寄存（Return internal error register）
END_FUNCTION_BLOCK
